(* IEC 61131-3 sources: Industry-PLC-LLM/data/PLCBEAD_repo/PLCBEAD_PLCEmbed-main/PLC-BEAD/Source/PLC_Programs (part 13) *)

(* ---- TN_SC_AREA_RESTORE.ST ---- *)
TYPE
  bya_TN_CHAR:       	ARRAY [0..1919] OF BYTE;
  bya_TN_BACKUP:     	ARRAY [0..1919] OF BYTE;
  bya_TN_COLOR:      	ARRAY [0..1919] OF BYTE;
  bya_TN_Line_Update:	ARRAY [0..23]   OF BOOL;

  us_TN_SCREEN :
  STRUCT
		bya_CHAR:			bya_TN_CHAR;
		bya_COLOR:			bya_TN_COLOR;
		bya_BACKUP:			bya_TN_BACKUP;
		bya_Line_Update:	bya_TN_Line_Update;

		by_Input_Exten_Code:    BYTE;
		by_Input_ASCII_Code:    BYTE;
		bo_Input_ASCII_IsNum:   BOOL;
		in_Page_Number:        	INT;                (* aktive Seiten-Nr.              *)
		in_Cursor_X:           	INT;                (* Cursor X-Position              *)
		in_Cursor_Y:           	INT;                (* Cursor Y-Position              *)
		in_EOS_Offset:         	INT;                (* End of String Offset           *)
		by_Clear_Screen_Attr:  	BYTE;               (* Clear-Screen Attr              *)
		bo_Clear_Screen:       	BOOL;               (* Clear-Screen ausl�sen          *)
		bo_Modal_Dialog:       	BOOL;               (* Modaler Dialog ist aktiv       *)
		bo_Menue_Bar_Dialog:   	BOOL;               (* Menue Dialog ist aktiv         *)

  END_STRUCT;
END_TYPE

FUNCTION TN_SC_XY2_ERROR:BOOL

	VAR_INPUT
		X1 :	INT;
		Y1 :	INT;
		X2 :	INT;
		Y2 :	INT;
	END_VAR

	TN_SC_XY2_ERROR := Y1 < 0 OR X1 < 0 OR Y2 < 0 OR X2 < 0 OR Y1 > 23 OR X1 > 79 OR Y2 > 23 OR X2 > 79;

END_FUNCTION

FUNCTION _BYTE_TO_INT:INT
	VAR_INPUT
		IN :	BYTE;
	END_VAR

	_BYTE_TO_INT := USINT_TO_INT(BYTE_TO_USINT(IN));
END_FUNCTION

FUNCTION_BLOCK TN_SC_AREA_RESTORE_Block

  VAR
    in_Offset_1 :	INT;
    in_Offset_2 :	INT;
    in_Y :	INT;
    in_X :	INT;
    in_Y1 :	INT;
    in_X1 :	INT;
    in_Y2 :	INT;
    in_X2 :	INT;
  END_VAR

  VAR_IN_OUT
    Xus_TN_SCREEN :	us_TN_SCREEN;
  END_VAR

  IF Xus_TN_SCREEN.bya_BACKUP[0] > BYTE#00 THEN

    in_X1 := _BYTE_TO_INT(Xus_TN_SCREEN.bya_BACKUP[1]);
    in_Y1 := _BYTE_TO_INT(Xus_TN_SCREEN.bya_BACKUP[2]);
    in_X2 := _BYTE_TO_INT(Xus_TN_SCREEN.bya_BACKUP[3]);
    in_Y2 := _BYTE_TO_INT(Xus_TN_SCREEN.bya_BACKUP[4]);

    IF TN_SC_XY2_ERROR(in_X1,in_Y1,in_X2,in_Y2) THEN RETURN; END_IF;
    in_Offset_2 := 5;

    FOR in_Y := in_Y1 TO in_Y2 DO

      Xus_TN_SCREEN.bya_Line_Update[in_Y] := TRUE;
      in_Offset_1 := (in_Y * 80) + in_X1;

      FOR in_X := in_X1 TO in_X2 DO

        Xus_TN_SCREEN.bya_CHAR[in_Offset_1] := Xus_TN_SCREEN.bya_BACKUP[in_Offset_2];
        in_Offset_2 := in_Offset_2 + INT#01;

        Xus_TN_SCREEN.bya_COLOR[in_Offset_1] := Xus_TN_SCREEN.bya_BACKUP[in_Offset_2];
        in_Offset_2 := in_Offset_2 + INT#01;
        in_Offset_1 := in_Offset_1 + INT#01;

      END_FOR;

    END_FOR;

    Xus_TN_SCREEN.bya_BACKUP[0] := BYTE#00;
  END_IF;

END_FUNCTION_BLOCK

PROGRAM program0
	VAR
		Xus_TN_SCREEN :	us_TN_SCREEN;

		func_block : TN_SC_AREA_RESTORE_Block;
	END_VAR
	func_block.Xus_TN_SCREEN := Xus_TN_SCREEN;

	func_block();
	Xus_TN_SCREEN  := func_block.Xus_TN_SCREEN;
END_PROGRAM

CONFIGURATION Config0
	RESOURCE Res0 ON PLC
		TASK task0(INTERVAL := T#20ms,PRIORITY := 0);
		PROGRAM instance0 WITH task0 : program0;
	END_RESOURCE
END_CONFIGURATION

(* ---- TN_SC_AREA_SAVE.ST ---- *)
TYPE
  bya_TN_CHAR:       	ARRAY [0..1919] OF BYTE;
  bya_TN_BACKUP:     	ARRAY [0..1919] OF BYTE;
  bya_TN_COLOR:      	ARRAY [0..1919] OF BYTE;
  bya_TN_Line_Update:	ARRAY [0..23]   OF BOOL;

  us_TN_SCREEN :
  STRUCT
		bya_CHAR:			bya_TN_CHAR;
		bya_COLOR:			bya_TN_COLOR;
		bya_BACKUP:			bya_TN_BACKUP;
		bya_Line_Update:	bya_TN_Line_Update;

		by_Input_Exten_Code:    BYTE;
		by_Input_ASCII_Code:    BYTE;
		bo_Input_ASCII_IsNum:   BOOL;
		in_Page_Number:        	INT;                (* aktive Seiten-Nr.              *)
		in_Cursor_X:           	INT;                (* Cursor X-Position              *)
		in_Cursor_Y:           	INT;                (* Cursor Y-Position              *)
		in_EOS_Offset:         	INT;                (* End of String Offset           *)
		by_Clear_Screen_Attr:  	BYTE;               (* Clear-Screen Attr              *)
		bo_Clear_Screen:       	BOOL;               (* Clear-Screen ausl�sen          *)
		bo_Modal_Dialog:       	BOOL;               (* Modaler Dialog ist aktiv       *)
		bo_Menue_Bar_Dialog:   	BOOL;               (* Menue Dialog ist aktiv         *)

  END_STRUCT;
END_TYPE

FUNCTION TN_SC_XY2_ERROR:BOOL

	VAR_INPUT
		X1 :	INT;
		Y1 :	INT;
		X2 :	INT;
		Y2 :	INT;
	END_VAR

	TN_SC_XY2_ERROR := Y1 < 0 OR X1 < 0 OR Y2 < 0 OR X2 < 0 OR Y1 > 23 OR X1 > 79 OR Y2 > 23 OR X2 > 79;

END_FUNCTION

FUNCTION_BLOCK TN_SC_AREA_SAVE_Block

	VAR
		in_Offset_1 :	INT;
		in_Offset_2 :	INT;
		in_Y :	INT;
		in_X :	INT;
	END_VAR

	VAR_INPUT
		Iin_Y1 :	INT;
		Iin_X1 :	INT;
		Iin_Y2 :	INT;
		Iin_X2 :	INT;
	END_VAR

	VAR_IN_OUT
		Xus_TN_SCREEN :	us_TN_SCREEN;
	END_VAR

	IF TN_SC_XY2_ERROR(Iin_X1,Iin_Y1,Iin_X2,Iin_Y2) THEN RETURN; END_IF;

	Xus_TN_SCREEN.bya_BACKUP[0] := BYTE#1;
	Xus_TN_SCREEN.bya_BACKUP[1] := INT_TO_BYTE(Iin_X1);
	Xus_TN_SCREEN.bya_BACKUP[2] := INT_TO_BYTE(Iin_Y1);
	Xus_TN_SCREEN.bya_BACKUP[3] := INT_TO_BYTE(Iin_X2);
	Xus_TN_SCREEN.bya_BACKUP[4] := INT_TO_BYTE(Iin_Y2);

	in_Offset_2 := 5;
	FOR in_Y := Iin_Y1 TO Iin_Y2 DO

	in_Offset_1 := (in_Y * 80) + Iin_X1;
	FOR in_X := Iin_X1 TO Iin_X2 DO

		Xus_TN_SCREEN.bya_BACKUP[in_Offset_2] := Xus_TN_SCREEN.bya_CHAR[in_Offset_1];
		in_Offset_2 := in_Offset_2 + INT#01;
		Xus_TN_SCREEN.bya_BACKUP[in_Offset_2] := Xus_TN_SCREEN.bya_COLOR[in_Offset_1];
		in_Offset_2 := in_Offset_2 + INT#01;
		in_Offset_1 := in_Offset_1 + INT#01;

	END_FOR;
	END_FOR;

END_FUNCTION_BLOCK

PROGRAM program0
	VAR
		Iin_Y1 :	INT;
		Iin_X1 :	INT;
		Iin_Y2 :	INT;
		Iin_X2 :	INT;
		Xus_TN_SCREEN :	us_TN_SCREEN;

		func_block : TN_SC_AREA_SAVE_Block;
	END_VAR
	func_block.Iin_X1 := Iin_X1;
	func_block.Iin_Y1 := Iin_Y1;
	func_block.Iin_X2 := Iin_X2;
	func_block.Iin_Y2 := Iin_Y2;
	func_block.Xus_TN_SCREEN := Xus_TN_SCREEN;

	func_block();
	Xus_TN_SCREEN  := func_block.Xus_TN_SCREEN;
END_PROGRAM

CONFIGURATION Config0
	RESOURCE Res0 ON PLC
		TASK task0(INTERVAL := T#20ms,PRIORITY := 0);
		PROGRAM instance0 WITH task0 : program0;
	END_RESOURCE
END_CONFIGURATION

(* ---- TN_SC_BOX.ST ---- *)
TYPE
  bya_TN_CHAR:       	ARRAY [0..1919] OF BYTE;
  bya_TN_BACKUP:     	ARRAY [0..1919] OF BYTE;
  bya_TN_COLOR:      	ARRAY [0..1919] OF BYTE;
  bya_TN_Line_Update:	ARRAY [0..23]   OF BOOL;

  us_TN_SCREEN :
  STRUCT
		bya_CHAR:			bya_TN_CHAR;
		bya_COLOR:			bya_TN_COLOR;
		bya_BACKUP:			bya_TN_BACKUP;
		bya_Line_Update:	bya_TN_Line_Update;

		by_Input_Exten_Code:    BYTE;
		by_Input_ASCII_Code:    BYTE;
		bo_Input_ASCII_IsNum:   BOOL;
		in_Page_Number:        	INT;                (* aktive Seiten-Nr.              *)
		in_Cursor_X:           	INT;                (* Cursor X-Position              *)
		in_Cursor_Y:           	INT;                (* Cursor Y-Position              *)
		in_EOS_Offset:         	INT;                (* End of String Offset           *)
		by_Clear_Screen_Attr:  	BYTE;               (* Clear-Screen Attr              *)
		bo_Clear_Screen:       	BOOL;               (* Clear-Screen ausl�sen          *)
		bo_Modal_Dialog:       	BOOL;               (* Modaler Dialog ist aktiv       *)
		bo_Menue_Bar_Dialog:   	BOOL;               (* Menue Dialog ist aktiv         *)

  END_STRUCT;
END_TYPE

FUNCTION TN_SC_XY2_ERROR:BOOL

	VAR_INPUT
		X1 :	INT;
		Y1 :	INT;
		X2 :	INT;
		Y2 :	INT;
	END_VAR

	TN_SC_XY2_ERROR := Y1 < 0 OR X1 < 0 OR Y2 < 0 OR X2 < 0 OR Y1 > 23 OR X1 > 79 OR Y2 > 23 OR X2 > 79;

END_FUNCTION

FUNCTION_BLOCK TN_SC_FILL_Block

	VAR
		in_X :	INT;
		in_Y :	INT;
		in_Offset :	INT;
	END_VAR

	VAR_INPUT
		Iin_Y1 :	INT;
		Iin_X1 :	INT;
		Iin_Y2 :	INT;
		Iin_X2 :	INT;
		Iby_CHAR :	BYTE;
		Iby_Attr :	BYTE;
	END_VAR

	VAR_IN_OUT
		Xus_TN_SCREEN :	us_TN_SCREEN;
	END_VAR

	IF TN_SC_XY2_ERROR(Iin_X1,Iin_Y1,Iin_X2,Iin_Y2) THEN RETURN; END_IF;

	FOR in_Y := Iin_Y1 TO Iin_Y2 DO
	Xus_TN_SCREEN.bya_Line_Update[in_Y] := TRUE;
	in_Offset := (in_Y * 80) + Iin_X1;
	FOR in_X := Iin_X1 TO Iin_X2 DO
		Xus_TN_SCREEN.bya_CHAR[in_Offset]  := Iby_CHAR;
		Xus_TN_SCREEN.bya_COLOR[in_Offset] := Iby_Attr;
		in_Offset := in_Offset + 1;
	END_FOR;
	END_FOR;

END_FUNCTION_BLOCK

FUNCTION_BLOCK TN_SC_BOX_Block

  VAR
    FB_TN_SC_FILL :	TN_SC_FILL_Block;
  END_VAR

  VAR
    by_BorderChar_L_T :	BYTE;
    by_BorderChar_T :	BYTE;
    by_BorderChar_B :	BYTE;
    by_BorderChar_R_T :	BYTE;
    by_BorderChar_L :	BYTE;
    by_BorderChar_R :	BYTE;
    by_BorderChar_L_B :	BYTE;
    by_BorderChar_R_B :	BYTE;
    in_Y :	INT;
    in_X :	INT;
    in_Border_Offset :	INT;
    in_Offset_1 :	INT;
    in_Offset_2 :	INT;
  END_VAR

  VAR_INPUT
    Iin_Y1 :	INT;
    Iin_X1 :	INT;
    Iin_Y2 :	INT;
    Iin_X2 :	INT;
    Iby_FILL :	BYTE;
    Iby_ATTR :	BYTE;
    Iin_BORDER :	INT;
  END_VAR

  VAR_IN_OUT
    Xus_TN_SCREEN :	us_TN_SCREEN;
  END_VAR

  IF TN_SC_XY2_ERROR(Iin_X1,Iin_Y1,Iin_X2,Iin_Y2) THEN RETURN; END_IF;

  CASE Iin_Border OF
  0:
    in_Border_Offset := 0;

  1:
    by_BorderChar_L_T := BYTE#218;
    by_BorderChar_T   := BYTE#196;
    by_BorderChar_R_T := BYTE#191;
    by_BorderChar_L   := BYTE#179;
    by_BorderChar_R   := BYTE#179;
    by_BorderChar_B   := BYTE#196;
    by_BorderChar_L_B := BYTE#217;
    by_BorderChar_R_B := BYTE#192;
    in_Border_Offset  := 1;

  2:
    by_BorderChar_L_T := BYTE#201;
    by_BorderChar_T   := BYTE#205;
    by_BorderChar_R_T := BYTE#187;
    by_BorderChar_L   := BYTE#186;
    by_BorderChar_R   := BYTE#186;
    by_BorderChar_B   := BYTE#205;
    by_BorderChar_L_B := BYTE#188;
    by_BorderChar_R_B := BYTE#200;
    in_Border_Offset  := 1;

  ELSE
    by_BorderChar_L_T := BYTE#32;
    by_BorderChar_T   := BYTE#32;
    by_BorderChar_R_T := BYTE#32;
    by_BorderChar_L   := BYTE#32;
    by_BorderChar_R   := BYTE#32;
    by_BorderChar_B   := BYTE#32;
    by_BorderChar_L_B := BYTE#32;
    by_BorderChar_R_B := BYTE#32;
    in_Border_Offset  := 1;

  END_CASE;

  IF Iby_FILL > BYTE#0 THEN

    FB_TN_SC_FILL.Iin_Y1			:= Iin_Y1 + in_Border_Offset;
    FB_TN_SC_FILL.Iin_X1			:= Iin_X1 + in_Border_Offset;
    FB_TN_SC_FILL.Iin_Y2			:= Iin_Y2 - in_Border_Offset;
    FB_TN_SC_FILL.Iin_X2			:= Iin_X2 - in_Border_Offset;
    FB_TN_SC_FILL.Iby_CHAR		:= Iby_FILL;
    FB_TN_SC_FILL.Iby_Attr		:= Iby_ATTR;
    FB_TN_SC_FILL.Xus_TN_SCREEN := Xus_TN_SCREEN;
    FB_TN_SC_FILL();
    Xus_TN_SCREEN := FB_TN_SC_FILL.Xus_TN_SCREEN;

  END_IF;

  IF Iin_BORDER = 0 THEN RETURN; END_IF;

  in_Offset_1 := (Iin_Y1 * 80) + Iin_X1;
  in_Offset_2 := (Iin_Y1 * 80) + Iin_X2;

  FOR in_Y := Iin_Y1 TO Iin_Y2 DO

    Xus_TN_SCREEN.bya_Line_Update[in_Y] := TRUE;

    Xus_TN_SCREEN.bya_CHAR[in_Offset_1]  := by_BorderChar_L;
    Xus_TN_SCREEN.bya_COLOR[in_Offset_1] := Iby_Attr;

    Xus_TN_SCREEN.bya_CHAR[in_Offset_2]  := by_BorderChar_R;
    Xus_TN_SCREEN.bya_COLOR[in_Offset_2] := Iby_Attr;

    in_Offset_1 := in_Offset_1 + 80;
    in_Offset_2 := in_Offset_2 + 80;

  END_FOR;

  in_Offset_1 := (Iin_Y1 * 80) + Iin_X1;
  in_Offset_2 := (Iin_Y2 * 80) + Iin_X1;

  FOR in_X := Iin_X1 TO Iin_X2 DO

    Xus_TN_SCREEN.bya_CHAR[in_Offset_1]  := by_BorderChar_T;
    Xus_TN_SCREEN.bya_COLOR[in_Offset_1] := Iby_Attr;

    Xus_TN_SCREEN.bya_CHAR[in_Offset_2]  := by_BorderChar_B;
    Xus_TN_SCREEN.bya_COLOR[in_Offset_2] := Iby_Attr;

    in_Offset_1 := in_Offset_1 + INT#1;
    in_Offset_2 := in_Offset_2 + INT#1;

  END_FOR;

  in_Offset_1 := (Iin_Y1 * 80) + Iin_X1;
  Xus_TN_SCREEN.bya_CHAR[in_Offset_1]  := by_BorderChar_L_T;
  Xus_TN_SCREEN.bya_COLOR[in_Offset_1] := Iby_Attr;

  in_Offset_1 := (Iin_Y1 * 80) + Iin_X2;
  Xus_TN_SCREEN.bya_CHAR[in_Offset_1]  := by_BorderChar_R_T;
  Xus_TN_SCREEN.bya_COLOR[in_Offset_1] := Iby_Attr;

  in_Offset_1 := (Iin_Y2 * 80) + Iin_X1;
  Xus_TN_SCREEN.bya_CHAR[in_Offset_1]  := by_BorderChar_R_B;
  Xus_TN_SCREEN.bya_COLOR[in_Offset_1] := Iby_Attr;

  in_Offset_1 := (Iin_Y2 * 80) + Iin_X2;
  Xus_TN_SCREEN.bya_CHAR[in_Offset_1]  := by_BorderChar_L_B;
  Xus_TN_SCREEN.bya_COLOR[in_Offset_1] := Iby_Attr;

END_FUNCTION_BLOCK

PROGRAM program0
	VAR
		Iin_Y1 :	INT;
    Iin_X1 :	INT;
    Iin_Y2 :	INT;
    Iin_X2 :	INT;
    Iby_FILL :	BYTE;
    Iby_ATTR :	BYTE;
    Iin_BORDER :	INT;
		Xus_TN_SCREEN :	us_TN_SCREEN;

		func_block : TN_SC_BOX_Block;
	END_VAR
  func_block.Iin_X1 := Iin_X1;
  func_block.Iin_Y1 := Iin_Y1;
  func_block.Iin_X2 := Iin_X2;
  func_block.Iin_Y2 := Iin_Y2;
  func_block.Iby_FILL := Iby_FILL;
  func_block.Iby_ATTR := Iby_ATTR;
  func_block.Iin_BORDER := Iin_BORDER;
  func_block.Xus_TN_SCREEN := Xus_TN_SCREEN;

	func_block();
	Xus_TN_SCREEN  := func_block.Xus_TN_SCREEN;
END_PROGRAM

CONFIGURATION Config0
	RESOURCE Res0 ON PLC
		TASK task0(INTERVAL := T#20ms,PRIORITY := 0);
		PROGRAM instance0 WITH task0 : program0;
	END_RESOURCE
END_CONFIGURATION

(* ---- TN_SC_FILL.ST ---- *)
TYPE
  bya_TN_CHAR:       	ARRAY [0..1919] OF BYTE;
  bya_TN_BACKUP:     	ARRAY [0..1919] OF BYTE;
  bya_TN_COLOR:      	ARRAY [0..1919] OF BYTE;
  bya_TN_Line_Update:	ARRAY [0..23]   OF BOOL;

  us_TN_SCREEN :
  STRUCT
		bya_CHAR:			bya_TN_CHAR;
		bya_COLOR:			bya_TN_COLOR;
		bya_BACKUP:			bya_TN_BACKUP;
		bya_Line_Update:	bya_TN_Line_Update;

		by_Input_Exten_Code:    BYTE;
		by_Input_ASCII_Code:    BYTE;
		bo_Input_ASCII_IsNum:   BOOL;
		in_Page_Number:        	INT;                (* aktive Seiten-Nr.              *)
		in_Cursor_X:           	INT;                (* Cursor X-Position              *)
		in_Cursor_Y:           	INT;                (* Cursor Y-Position              *)
		in_EOS_Offset:         	INT;                (* End of String Offset           *)
		by_Clear_Screen_Attr:  	BYTE;               (* Clear-Screen Attr              *)
		bo_Clear_Screen:       	BOOL;               (* Clear-Screen ausl�sen          *)
		bo_Modal_Dialog:       	BOOL;               (* Modaler Dialog ist aktiv       *)
		bo_Menue_Bar_Dialog:   	BOOL;               (* Menue Dialog ist aktiv         *)

  END_STRUCT;
END_TYPE

FUNCTION TN_SC_XY2_ERROR:BOOL

	VAR_INPUT
		X1 :	INT;
		Y1 :	INT;
		X2 :	INT;
		Y2 :	INT;
	END_VAR

	TN_SC_XY2_ERROR := Y1 < 0 OR X1 < 0 OR Y2 < 0 OR X2 < 0 OR Y1 > 23 OR X1 > 79 OR Y2 > 23 OR X2 > 79;

END_FUNCTION

FUNCTION_BLOCK TN_SC_FILL_Block

	VAR
		in_X :	INT;
		in_Y :	INT;
		in_Offset :	INT;
	END_VAR

	VAR_INPUT
		Iin_Y1 :	INT;
		Iin_X1 :	INT;
		Iin_Y2 :	INT;
		Iin_X2 :	INT;
		Iby_CHAR :	BYTE;
		Iby_Attr :	BYTE;
	END_VAR

	VAR_IN_OUT
		Xus_TN_SCREEN :	us_TN_SCREEN;
	END_VAR

	IF TN_SC_XY2_ERROR(Iin_X1,Iin_Y1,Iin_X2,Iin_Y2) THEN RETURN; END_IF;

	FOR in_Y := Iin_Y1 TO Iin_Y2 DO
	Xus_TN_SCREEN.bya_Line_Update[in_Y] := TRUE;
	in_Offset := (in_Y * 80) + Iin_X1;
	FOR in_X := Iin_X1 TO Iin_X2 DO
		Xus_TN_SCREEN.bya_CHAR[in_Offset]  := Iby_CHAR;
		Xus_TN_SCREEN.bya_COLOR[in_Offset] := Iby_Attr;
		in_Offset := in_Offset + 1;
	END_FOR;
	END_FOR;

END_FUNCTION_BLOCK

PROGRAM program0
	VAR
		Iin_Y1 :	INT;
		Iin_X1 :	INT;
		Iin_Y2 :	INT;
		Iin_X2 :	INT;
		Iby_CHAR :	BYTE;
		Iby_Attr :	BYTE;
		Xus_TN_SCREEN :	us_TN_SCREEN;

		func_block : TN_SC_FILL_Block;
	END_VAR
	func_block.Iin_X1 := Iin_X1;
	func_block.Iin_Y1 := Iin_Y1;
  	func_block.Iin_X2 := Iin_X2;
	func_block.Iin_Y2 := Iin_Y2;
  	func_block.Iby_CHAR := Iby_CHAR;
	func_block.Iby_Attr := Iby_Attr;
	func_block.Xus_TN_SCREEN := Xus_TN_SCREEN;

	func_block();
	Xus_TN_SCREEN  := func_block.Xus_TN_SCREEN;
END_PROGRAM

CONFIGURATION Config0
	RESOURCE Res0 ON PLC
		TASK task0(INTERVAL := T#20ms,PRIORITY := 0);
		PROGRAM instance0 WITH task0 : program0;
	END_RESOURCE
END_CONFIGURATION

(* ---- TN_SC_LINE.ST ---- *)
TYPE
  bya_TN_CHAR:       	ARRAY [0..1919] OF BYTE;
  bya_TN_BACKUP:     	ARRAY [0..1919] OF BYTE;
  bya_TN_COLOR:      	ARRAY [0..1919] OF BYTE;
  bya_TN_Line_Update:	ARRAY [0..23]   OF BOOL;

  us_TN_SCREEN :
  STRUCT
		bya_CHAR:			bya_TN_CHAR;
		bya_COLOR:			bya_TN_COLOR;
		bya_BACKUP:			bya_TN_BACKUP;
		bya_Line_Update:	bya_TN_Line_Update;

		by_Input_Exten_Code:    BYTE;
		by_Input_ASCII_Code:    BYTE;
		bo_Input_ASCII_IsNum:   BOOL;
		in_Page_Number:        	INT;                (* aktive Seiten-Nr.              *)
		in_Cursor_X:           	INT;                (* Cursor X-Position              *)
		in_Cursor_Y:           	INT;                (* Cursor Y-Position              *)
		in_EOS_Offset:         	INT;                (* End of String Offset           *)
		by_Clear_Screen_Attr:  	BYTE;               (* Clear-Screen Attr              *)
		bo_Clear_Screen:       	BOOL;               (* Clear-Screen ausl�sen          *)
		bo_Modal_Dialog:       	BOOL;               (* Modaler Dialog ist aktiv       *)
		bo_Menue_Bar_Dialog:   	BOOL;               (* Menue Dialog ist aktiv         *)

  END_STRUCT;
END_TYPE

FUNCTION TN_SC_XY2_ERROR:BOOL

	VAR_INPUT
		X1 :	INT;
		Y1 :	INT;
		X2 :	INT;
		Y2 :	INT;
	END_VAR

	TN_SC_XY2_ERROR := Y1 < 0 OR X1 < 0 OR Y2 < 0 OR X2 < 0 OR Y1 > 23 OR X1 > 79 OR Y2 > 23 OR X2 > 79;

END_FUNCTION

FUNCTION_BLOCK TN_SC_LINE_Block

  VAR
    by_Connect_Left_Char :	BYTE;
    by_Connect_Right_Char :	BYTE;
    by_Connect_Top_Char :	BYTE;
    by_Connect_Bottom_Char :	BYTE;
    by_Connect_Cruz_Char :	BYTE;
    by_Vertikal_Line_Char :	BYTE;
    by_Horzontal_Line_Char :	BYTE;
    by_old_Char :	BYTE;
    in_Offset_1 :	INT;
    in_ROW_Index :	INT;
    in_COL_Index :	INT;
    by_Char :	BYTE;
  END_VAR

  VAR_INPUT
    Iin_X1 :	INT;
    Iin_Y1 :	INT;
    Iin_X2 :	INT;
    Iin_Y2 :	INT;
    Iby_ATTR :	BYTE;
    Iby_BORDER :	BYTE;
  END_VAR

  VAR_IN_OUT
    Xus_TN_SCREEN :	us_TN_SCREEN;
  END_VAR

  IF TN_SC_XY2_ERROR(Iin_X1,Iin_Y1,Iin_X2,Iin_Y2) THEN RETURN; END_IF;

  IF Iby_Border = BYTE#01 THEN

    by_Connect_Top_Char    := BYTE#16#C2;
    by_Connect_Bottom_Char := BYTE#16#C1;
    by_Connect_Left_Char   := BYTE#16#C3;
    by_Connect_Right_Char  := BYTE#16#B4;
    by_Horzontal_Line_Char := BYTE#16#C4;
    by_Vertikal_Line_Char  := BYTE#16#B3;
    by_Connect_Cruz_Char   := BYTE#16#C5;

  ELSIF Iby_Border = BYTE#02 THEN

    by_Connect_Top_Char    := BYTE#16#CB;
    by_Connect_Bottom_Char := BYTE#16#CA;
    by_Connect_Left_Char   := BYTE#16#CC;
    by_Connect_Right_Char  := BYTE#16#B9;
    by_Horzontal_Line_Char := BYTE#16#CD;
    by_Vertikal_Line_Char  := BYTE#16#BA;
    by_Connect_Cruz_Char   := BYTE#16#CE;

  ELSE
    by_Connect_Top_Char    := Iby_Border;
    by_Connect_Bottom_Char := Iby_Border;
    by_Connect_Left_Char   := Iby_Border;
    by_Connect_Right_Char  := Iby_Border;
    by_Horzontal_Line_Char := Iby_Border;
    by_Vertikal_Line_Char  := Iby_Border;
    by_Connect_Cruz_Char   := Iby_Border;

  END_IF;

  IF Iin_X1 = Iin_X2 THEN

    in_Offset_1 := (Iin_Y1 * 80) + Iin_X1;

    FOR in_ROW_Index := Iin_Y1 TO Iin_Y2 DO

      by_old_Char := Xus_TN_SCREEN.bya_CHAR[in_Offset_1];

      by_Char := by_Vertikal_Line_Char;

      IF by_old_Char = by_Horzontal_Line_Char THEN

        IF in_ROW_Index = Iin_Y1 THEN
          by_Char := by_Connect_Top_Char;

        ELSIF in_ROW_Index = Iin_Y2 THEN
          by_Char := by_Connect_Bottom_Char;

        ELSE
          by_Char := by_Connect_Cruz_Char;
        END_IF;

      END_IF;

      Xus_TN_SCREEN.bya_Line_Update[in_ROW_Index] := TRUE;

      Xus_TN_SCREEN.bya_CHAR[in_Offset_1]  := by_Char;
      Xus_TN_SCREEN.bya_COLOR[in_Offset_1] := Iby_Attr;

      in_Offset_1 := in_Offset_1 + 80;

    END_FOR;

  ELSIF Iin_Y1 = Iin_Y2 THEN

    Xus_TN_SCREEN.bya_Line_Update[Iin_Y1] := TRUE;

    in_Offset_1 := (Iin_Y1 * 80) + Iin_X1;

    FOR in_COL_Index := Iin_X1 TO Iin_X2 DO

      by_old_Char := Xus_TN_SCREEN.bya_CHAR[in_Offset_1];

      by_Char := by_Horzontal_Line_Char;

      IF by_old_Char = by_Vertikal_Line_Char THEN

        IF in_COL_Index = Iin_X1 THEN
          by_Char := by_Connect_Left_Char;

        ELSIF in_COL_Index = Iin_X2 THEN
          by_Char := by_Connect_Right_Char;

        ELSE
          by_Char := by_Connect_Cruz_Char;
        END_IF;

      END_IF;

      Xus_TN_SCREEN.bya_CHAR[in_Offset_1]  := by_Char;
      Xus_TN_SCREEN.bya_COLOR[in_Offset_1] := Iby_Attr;

      in_Offset_1 := in_Offset_1 + 1;

    END_FOR;
  END_IF;

END_FUNCTION_BLOCK

PROGRAM program0
	VAR
    Iin_X1 :	INT;
    Iin_Y1 :	INT;
    Iin_X2 :	INT;
    Iin_Y2 :	INT;
    Iby_ATTR :	BYTE;
    Iby_BORDER :	BYTE;
    Xus_TN_SCREEN :	us_TN_SCREEN;

    func_block : TN_SC_LINE_Block;
	END_VAR
	func_block.Iin_X1 := Iin_X1;
	func_block.Iin_Y1 := Iin_Y1;
  func_block.Iin_X2 := Iin_X2;
	func_block.Iin_Y2 := Iin_Y2;
  func_block.Iby_ATTR := Iby_ATTR;
	func_block.Iby_BORDER := Iby_BORDER;
	func_block.Xus_TN_SCREEN := Xus_TN_SCREEN;

	func_block();
	Xus_TN_SCREEN  := func_block.Xus_TN_SCREEN;
END_PROGRAM

CONFIGURATION Config0
	RESOURCE Res0 ON PLC
		TASK task0(INTERVAL := T#20ms,PRIORITY := 0);
		PROGRAM instance0 WITH task0 : program0;
	END_RESOURCE
END_CONFIGURATION

(* ---- TN_SC_READ_ATTR.ST ---- *)
TYPE
  bya_TN_CHAR:       	ARRAY [0..1919] OF BYTE;
  bya_TN_BACKUP:     	ARRAY [0..1919] OF BYTE;
  bya_TN_COLOR:      	ARRAY [0..1919] OF BYTE;
  bya_TN_Line_Update:	ARRAY [0..23]   OF BOOL;

  us_TN_SCREEN :
  STRUCT
		bya_CHAR:			bya_TN_CHAR;
		bya_COLOR:			bya_TN_COLOR;
		bya_BACKUP:			bya_TN_BACKUP;
		bya_Line_Update:	bya_TN_Line_Update;

		by_Input_Exten_Code:    BYTE;
		by_Input_ASCII_Code:    BYTE;
		bo_Input_ASCII_IsNum:   BOOL;
		in_Page_Number:        	INT;                (* aktive Seiten-Nr.              *)
		in_Cursor_X:           	INT;                (* Cursor X-Position              *)
		in_Cursor_Y:           	INT;                (* Cursor Y-Position              *)
		in_EOS_Offset:         	INT;                (* End of String Offset           *)
		by_Clear_Screen_Attr:  	BYTE;               (* Clear-Screen Attr              *)
		bo_Clear_Screen:       	BOOL;               (* Clear-Screen ausl�sen          *)
		bo_Modal_Dialog:       	BOOL;               (* Modaler Dialog ist aktiv       *)
		bo_Menue_Bar_Dialog:   	BOOL;               (* Menue Dialog ist aktiv         *)

  END_STRUCT;
END_TYPE

FUNCTION TN_SC_XY_ERROR:BOOL

	VAR_INPUT
		X :	INT;
		Y :	INT;
	END_VAR

	TN_SC_XY_ERROR := Y < 0 OR X < 0 OR Y > 23 OR X > 79;

END_FUNCTION

FUNCTION_BLOCK TN_SC_READ_ATTR_Block

	VAR
		in_Offset :	INT;
	END_VAR

	VAR_INPUT
		Iin_Y :	INT;
		Iin_X :	INT;
	END_VAR

	VAR_OUTPUT
		Oby_ATTR :	BYTE;
	END_VAR

	VAR_IN_OUT
		Xus_TN_SCREEN :	us_TN_SCREEN;
	END_VAR

	IF TN_SC_XY_ERROR(Iin_X,Iin_Y) THEN RETURN; END_IF;
	in_Offset := (Iin_Y * 80) + Iin_X;
	Oby_ATTR := Xus_TN_SCREEN.bya_COLOR[in_Offset];

END_FUNCTION_BLOCK

PROGRAM program0
	VAR
		Iin_Y :	INT;
		Iin_X :	INT;
		Xus_TN_SCREEN :	us_TN_SCREEN;
		Oby_ATTR :	BYTE;

		func_block : TN_SC_READ_ATTR_Block;
	END_VAR
	func_block.Iin_Y := Iin_Y;
	func_block.Iin_X := Iin_X;
	func_block.Xus_TN_SCREEN := Xus_TN_SCREEN;

	func_block();
	Xus_TN_SCREEN  := func_block.Xus_TN_SCREEN;
	Oby_ATTR  := func_block.Oby_ATTR;
END_PROGRAM

CONFIGURATION Config0
	RESOURCE Res0 ON PLC
		TASK task0(INTERVAL := T#20ms,PRIORITY := 0);
		PROGRAM instance0 WITH task0 : program0;
	END_RESOURCE
END_CONFIGURATION

(* ---- TN_SC_READ_CHAR.ST ---- *)
TYPE
  bya_TN_CHAR:       	ARRAY [0..1919] OF BYTE;
  bya_TN_BACKUP:     	ARRAY [0..1919] OF BYTE;
  bya_TN_COLOR:      	ARRAY [0..1919] OF BYTE;
  bya_TN_Line_Update:	ARRAY [0..23]   OF BOOL;

  us_TN_SCREEN :
  STRUCT
		bya_CHAR:			bya_TN_CHAR;
		bya_COLOR:			bya_TN_COLOR;
		bya_BACKUP:			bya_TN_BACKUP;
		bya_Line_Update:	bya_TN_Line_Update;

		by_Input_Exten_Code:    BYTE;
		by_Input_ASCII_Code:    BYTE;
		bo_Input_ASCII_IsNum:   BOOL;
		in_Page_Number:        	INT;                (* aktive Seiten-Nr.              *)
		in_Cursor_X:           	INT;                (* Cursor X-Position              *)
		in_Cursor_Y:           	INT;                (* Cursor Y-Position              *)
		in_EOS_Offset:         	INT;                (* End of String Offset           *)
		by_Clear_Screen_Attr:  	BYTE;               (* Clear-Screen Attr              *)
		bo_Clear_Screen:       	BOOL;               (* Clear-Screen ausl�sen          *)
		bo_Modal_Dialog:       	BOOL;               (* Modaler Dialog ist aktiv       *)
		bo_Menue_Bar_Dialog:   	BOOL;               (* Menue Dialog ist aktiv         *)

  END_STRUCT;
END_TYPE

FUNCTION TN_SC_XY_ERROR:BOOL

	VAR_INPUT
		X :	INT;
		Y :	INT;
	END_VAR

	TN_SC_XY_ERROR := Y < 0 OR X < 0 OR Y > 23 OR X > 79;

END_FUNCTION

FUNCTION_BLOCK TN_SC_READ_CHAR_Block

	VAR
		in_Offset :	INT;
	END_VAR

	VAR_INPUT
		Iin_Y :	INT;
		Iin_X :	INT;
	END_VAR

	VAR_OUTPUT
		Oby_CHAR :	BYTE;
	END_VAR

	VAR_IN_OUT
		Xus_TN_SCREEN :	us_TN_SCREEN;
	END_VAR

	IF TN_SC_XY_ERROR(Iin_X,Iin_Y) THEN RETURN; END_IF;
	in_Offset := (Iin_Y * 80) + Iin_X;
	Oby_CHAR := Xus_TN_SCREEN.bya_CHAR[in_Offset];

END_FUNCTION_BLOCK

PROGRAM program0
	VAR
		Iin_Y :	INT;
		Iin_X :	INT;
		Xus_TN_SCREEN :	us_TN_SCREEN;
		Oby_CHAR :	BYTE;

		func_block : TN_SC_READ_CHAR_Block;
	END_VAR
	func_block.Iin_Y := Iin_Y;
	func_block.Iin_X := Iin_X;
	func_block.Xus_TN_SCREEN := Xus_TN_SCREEN;

	func_block();
	Xus_TN_SCREEN  := func_block.Xus_TN_SCREEN;
	Oby_CHAR  := func_block.Oby_CHAR;
END_PROGRAM

CONFIGURATION Config0
	RESOURCE Res0 ON PLC
		TASK task0(INTERVAL := T#20ms,PRIORITY := 0);
		PROGRAM instance0 WITH task0 : program0;
	END_RESOURCE
END_CONFIGURATION

(* ---- TN_SC_VIEWPORT.ST ---- *)
TYPE
  bya_TN_CHAR:       	ARRAY [0..1919] OF BYTE;
  bya_TN_BACKUP:     	ARRAY [0..1919] OF BYTE;
  bya_TN_COLOR:      	ARRAY [0..1919] OF BYTE;
  bya_TN_Line_Update:	ARRAY [0..23]   OF BOOL;

  us_TN_SCREEN :
  STRUCT
		bya_CHAR:			bya_TN_CHAR;
		bya_COLOR:			bya_TN_COLOR;
		bya_BACKUP:			bya_TN_BACKUP;
		bya_Line_Update:	bya_TN_Line_Update;

		by_Input_Exten_Code:    BYTE;
		by_Input_ASCII_Code:    BYTE;
		bo_Input_ASCII_IsNum:   BOOL;
		in_Page_Number:        	INT;                (* aktive Seiten-Nr.              *)
		in_Cursor_X:           	INT;                (* Cursor X-Position              *)
		in_Cursor_Y:           	INT;                (* Cursor Y-Position              *)
		in_EOS_Offset:         	INT;                (* End of String Offset           *)
		by_Clear_Screen_Attr:  	BYTE;               (* Clear-Screen Attr              *)
		bo_Clear_Screen:       	BOOL;               (* Clear-Screen ausl�sen          *)
		bo_Modal_Dialog:       	BOOL;               (* Modaler Dialog ist aktiv       *)
		bo_Menue_Bar_Dialog:   	BOOL;               (* Menue Dialog ist aktiv         *)

  END_STRUCT;
END_TYPE

FUNCTION_BLOCK TN_SC_VIEWPORT_Block

  VAR
    FB_TN_SC_WRITE :	TN_SC_WRITE;
    FB_FIX :	FIX;
    FB_TON :	TON;
  END_VAR

  VAR
    in_index :	INT;
    in_Color :	INT;
    by_Attr :	BYTE;
    in_count :	INT;
  END_VAR

  VAR_IN_OUT
    Xus_LOG_VIEWPORT :	us_LOG_VIEWPORT;
    Xus_LOG_CONTROL :	us_LOG_CONTROL_80;
    Xus_TN_SCREEN :	us_TN_SCREEN;
  END_VAR

  VAR_INPUT
    Iin_X :	INT;
    Iin_Y :	INT;
    Iin_Width :	INT;
    Idw_ATTR_1 :	DWORD;
    Idw_ATTR_2 :	DWORD;
    Iti_TIME :	TIME;
  END_VAR

  IF Xus_LOG_VIEWPORT.UPDATE AND FB_TON.Q THEN

    Xus_LOG_VIEWPORT.UPDATE := FALSE;

    FOR in_count := 1 TO Xus_LOG_VIEWPORT.COUNT DO

      in_index := Xus_LOG_VIEWPORT.LINE_ARRAY[in_count];

    in_Color := DWORD_TO_INT(Xus_LOG_CONTROL.MSG_OPTION[in_index] AND DWORD#2#1111);

      CASE in_Color OF
        0..3: by_Attr := BYTE_OF_DWORD(Idw_ATTR_1,INT_TO_BYTE(in_Color));
        4..7: by_Attr := BYTE_OF_DWORD(Idw_ATTR_2,INT_TO_BYTE(in_Color));
      ELSE
      by_Attr := BYTE_OF_DWORD(Idw_ATTR_1,BYTE#0);
      END_CASE;

      FB_FIX.str := Xus_LOG_CONTROL.MSG[in_index];
      FB_FIX.L   := Iin_Width;
      FB_FIX.C   := BYTE#32;
      FB_FIX.M   := INT#00;
      FB_FIX();

      FB_TN_SC_WRITE.Iin_Y			:= Iin_Y + in_count - INT#01;
      FB_TN_SC_WRITE.Iin_X			:= Iin_X;
      FB_TN_SC_WRITE.Iby_ATTR			:= by_Attr;
      FB_TN_SC_WRITE.Ist_STRING		:= FB_FIX.FIX;
      FB_TN_SC_WRITE.Xus_TN_SCREEN	:= Xus_TN_SCREEN;
      FB_TN_SC_WRITE();
      Xus_TN_SCREEN := FB_TN_SC_WRITE.Xus_TN_SCREEN;

    END_FOR;

    FB_TON.IN := FALSE;
    FB_TON.PT := Iti_TIME;
    FB_TON();

  END_IF;

  FB_TON.IN := TRUE;
  FB_TON.PT := Iti_TIME;
  FB_TON();

END_FUNCTION_BLOCK

PROGRAM program0
	VAR
		Xus_LOG_VIEWPORT :	us_LOG_VIEWPORT;
    Xus_LOG_CONTROL :	us_LOG_CONTROL_80;
    Xus_TN_SCREEN :	us_TN_SCREEN;
    Iin_X :	INT;
    Iin_Y :	INT;
    Iin_Width :	INT;
    Idw_ATTR_1 :	DWORD;
    Idw_ATTR_2 :	DWORD;
    Iti_TIME :	TIME;

		func_block : TN_SC_VIEWPORT_Block;
	END_VAR
	func_block.Xus_LOG_VIEWPORT := Xus_LOG_VIEWPORT;
	func_block.Xus_LOG_CONTROL := Xus_LOG_CONTROL;
	func_block.Xus_TN_SCREEN := Xus_TN_SCREEN;
	func_block.Iin_X := Iin_X;
  func_block.Iin_Y := Iin_Y;
	func_block.Iin_Width := Iin_Width;
	func_block.Idw_ATTR_1 := Idw_ATTR_1;
	func_block.Idw_ATTR_2 := Idw_ATTR_2;
  func_block.Iti_TIME := Iti_TIME;

	func_block();
	Xus_LOG_VIEWPORT  := func_block.Xus_LOG_VIEWPORT;
  Xus_LOG_CONTROL  := func_block.Xus_LOG_CONTROL;
  Xus_TN_SCREEN  := func_block.Xus_TN_SCREEN;
END_PROGRAM

CONFIGURATION Config0
	RESOURCE Res0 ON PLC
		TASK task0(INTERVAL := T#20ms,PRIORITY := 0);
		PROGRAM instance0 WITH task0 : program0;
	END_RESOURCE
END_CONFIGURATION

(* ---- TN_SC_WRITE.ST ---- *)
TYPE
  bya_TN_CHAR:       	ARRAY [0..1919] OF BYTE;
  bya_TN_BACKUP:     	ARRAY [0..1919] OF BYTE;
  bya_TN_COLOR:      	ARRAY [0..1919] OF BYTE;
  bya_TN_Line_Update:	ARRAY [0..23]   OF BOOL;

  us_TN_SCREEN :
  STRUCT
		bya_CHAR:			bya_TN_CHAR;
		bya_COLOR:			bya_TN_COLOR;
		bya_BACKUP:			bya_TN_BACKUP;
		bya_Line_Update:	bya_TN_Line_Update;

		by_Input_Exten_Code:    BYTE;
		by_Input_ASCII_Code:    BYTE;
		bo_Input_ASCII_IsNum:   BOOL;
		in_Page_Number:        	INT;                (* aktive Seiten-Nr.              *)
		in_Cursor_X:           	INT;                (* Cursor X-Position              *)
		in_Cursor_Y:           	INT;                (* Cursor Y-Position              *)
		in_EOS_Offset:         	INT;                (* End of String Offset           *)
		by_Clear_Screen_Attr:  	BYTE;               (* Clear-Screen Attr              *)
		bo_Clear_Screen:       	BOOL;               (* Clear-Screen ausl�sen          *)
		bo_Modal_Dialog:       	BOOL;               (* Modaler Dialog ist aktiv       *)
		bo_Menue_Bar_Dialog:   	BOOL;               (* Menue Dialog ist aktiv         *)

  END_STRUCT;
END_TYPE

FUNCTION TN_SC_XY_ERROR:BOOL

	VAR_INPUT
		X :	INT;
		Y :	INT;
	END_VAR

	TN_SC_XY_ERROR := Y < 0 OR X < 0 OR Y > 23 OR X > 79;

END_FUNCTION

FUNCTION_BLOCK TN_SC_WRITE_Block

	VAR
		CODE :	CODE;
	END_VAR

	VAR
		bo_Color :	BOOL;
		in_Offset :	INT;
		in_Char_Index :	INT;
		in_String_Length :	INT;
	END_VAR

	VAR_INPUT
		Iin_Y :	INT;
		Iin_X :	INT;
		Iby_ATTR :	BYTE;
		Ist_STRING :	STRING;
	END_VAR

	VAR_IN_OUT
		Xus_TN_SCREEN :	us_TN_SCREEN;
	END_VAR

	in_String_Length := LEN(Ist_STRING);
	IF TN_SC_XY_ERROR(Iin_X + in_String_Length - 1,Iin_Y) THEN RETURN; END_IF;
	Xus_TN_SCREEN.bya_Line_Update[Iin_Y] := TRUE;
	in_Offset := (Iin_Y * 80) + Iin_X;
	bo_Color := Iby_ATTR <> BYTE#00;

	FOR in_Char_Index := 1 TO in_String_Length DO

	IF bo_Color THEN Xus_TN_SCREEN.bya_COLOR[in_Offset] := Iby_ATTR; END_IF;

	CODE(STR:=Ist_STRING,POS:=in_Char_Index);
	Xus_TN_SCREEN.bya_CHAR[in_Offset] := CODE.CODE;
	in_Offset := in_Offset + INT#1;

	END_FOR;

	Xus_TN_SCREEN.in_EOS_Offset := in_Offset;

END_FUNCTION_BLOCK

PROGRAM program0
	VAR
		Iin_Y :	INT;
		Iin_X :	INT;
		Iby_ATTR :	BYTE;
		Ist_STRING :	STRING;
		Xus_TN_SCREEN :	us_TN_SCREEN;

		func_block : TN_SC_WRITE_Block;
	END_VAR
	func_block.Iin_Y := Iin_Y;
	func_block.Iin_X := Iin_X;
	func_block.Iby_ATTR := Iby_ATTR;
	func_block.Ist_STRING := Ist_STRING;
	func_block.Xus_TN_SCREEN := Xus_TN_SCREEN;

	func_block();
	Xus_TN_SCREEN  := func_block.Xus_TN_SCREEN;

END_PROGRAM

CONFIGURATION Config0
	RESOURCE Res0 ON PLC
		TASK task0(INTERVAL := T#20ms,PRIORITY := 0);
		PROGRAM instance0 WITH task0 : program0;
	END_RESOURCE
END_CONFIGURATION

(* ---- TN_SC_WRITE_ATTR.ST ---- *)
TYPE
  bya_TN_CHAR:       	ARRAY [0..1919] OF BYTE;
  bya_TN_BACKUP:     	ARRAY [0..1919] OF BYTE;
  bya_TN_COLOR:      	ARRAY [0..1919] OF BYTE;
  bya_TN_Line_Update:	ARRAY [0..23]   OF BOOL;

  us_TN_SCREEN :
  STRUCT
		bya_CHAR:			bya_TN_CHAR;
		bya_COLOR:			bya_TN_COLOR;
		bya_BACKUP:			bya_TN_BACKUP;
		bya_Line_Update:	bya_TN_Line_Update;

		by_Input_Exten_Code:    BYTE;
		by_Input_ASCII_Code:    BYTE;
		bo_Input_ASCII_IsNum:   BOOL;
		in_Page_Number:        	INT;                (* aktive Seiten-Nr.              *)
		in_Cursor_X:           	INT;                (* Cursor X-Position              *)
		in_Cursor_Y:           	INT;                (* Cursor Y-Position              *)
		in_EOS_Offset:         	INT;                (* End of String Offset           *)
		by_Clear_Screen_Attr:  	BYTE;               (* Clear-Screen Attr              *)
		bo_Clear_Screen:       	BOOL;               (* Clear-Screen ausl�sen          *)
		bo_Modal_Dialog:       	BOOL;               (* Modaler Dialog ist aktiv       *)
		bo_Menue_Bar_Dialog:   	BOOL;               (* Menue Dialog ist aktiv         *)

  END_STRUCT;
END_TYPE

FUNCTION TN_SC_XY_ERROR:BOOL

	VAR_INPUT
		X :	INT;
		Y :	INT;
	END_VAR

	TN_SC_XY_ERROR := Y < 0 OR X < 0 OR Y > 23 OR X > 79;

END_FUNCTION

FUNCTION_BLOCK TN_SC_WRITE_ATTR_Block

	VAR
		in_Offset :	INT;
	END_VAR

	VAR_INPUT
		Iin_Y :	INT;
		Iin_X :	INT;
		Iby_ATTR :	BYTE;
	END_VAR

	VAR_IN_OUT
		Xus_TN_SCREEN :	us_TN_SCREEN;
	END_VAR

	IF TN_SC_XY_ERROR(Iin_X,Iin_Y) THEN RETURN; END_IF;
	in_Offset := (Iin_Y * 80) + Iin_X;
	Xus_TN_SCREEN.bya_COLOR[in_Offset] := Iby_ATTR;

END_FUNCTION_BLOCK

PROGRAM program0
	VAR
		Iin_Y :	INT;
		Iin_X :	INT;
		Iby_ATTR :	BYTE;
		Xus_TN_SCREEN :	us_TN_SCREEN;

		func_block : TN_SC_WRITE_ATTR_Block;
	END_VAR
	func_block.Iin_Y := Iin_Y;
	func_block.Iin_X := Iin_X;
	func_block.Iby_ATTR := Iby_ATTR;
	func_block.Xus_TN_SCREEN := Xus_TN_SCREEN;

	func_block();
	Xus_TN_SCREEN  := func_block.Xus_TN_SCREEN;
END_PROGRAM

CONFIGURATION Config0
	RESOURCE Res0 ON PLC
		TASK task0(INTERVAL := T#20ms,PRIORITY := 0);
		PROGRAM instance0 WITH task0 : program0;
	END_RESOURCE
END_CONFIGURATION

(* ---- TN_SC_WRITE_C.ST ---- *)
TYPE
  bya_TN_CHAR:       	ARRAY [0..1919] OF BYTE;
  bya_TN_BACKUP:     	ARRAY [0..1919] OF BYTE;
  bya_TN_COLOR:      	ARRAY [0..1919] OF BYTE;
  bya_TN_Line_Update:	ARRAY [0..23]   OF BOOL;

  us_TN_SCREEN :
  STRUCT
		bya_CHAR:			bya_TN_CHAR;
		bya_COLOR:			bya_TN_COLOR;
		bya_BACKUP:			bya_TN_BACKUP;
		bya_Line_Update:	bya_TN_Line_Update;

		by_Input_Exten_Code:    BYTE;
		by_Input_ASCII_Code:    BYTE;
		bo_Input_ASCII_IsNum:   BOOL;
		in_Page_Number:        	INT;                (* aktive Seiten-Nr.              *)
		in_Cursor_X:           	INT;                (* Cursor X-Position              *)
		in_Cursor_Y:           	INT;                (* Cursor Y-Position              *)
		in_EOS_Offset:         	INT;                (* End of String Offset           *)
		by_Clear_Screen_Attr:  	BYTE;               (* Clear-Screen Attr              *)
		bo_Clear_Screen:       	BOOL;               (* Clear-Screen ausl�sen          *)
		bo_Modal_Dialog:       	BOOL;               (* Modaler Dialog ist aktiv       *)
		bo_Menue_Bar_Dialog:   	BOOL;               (* Menue Dialog ist aktiv         *)

  END_STRUCT;
END_TYPE

FUNCTION _BYTE_TO_INT:INT
	VAR_INPUT
		IN :	BYTE;
	END_VAR

	_BYTE_TO_INT := USINT_TO_INT(BYTE_TO_USINT(IN));
END_FUNCTION

FUNCTION_BLOCK CHR_TO_STRING_Block
	VAR_INPUT
		C :	BYTE;
	END_VAR

	VAR_OUTPUT
		CHR_TO_STRING :	STRING;
	END_VAR

	CHR_TO_STRING := BYTE_TO_STRING(C);

END_FUNCTION_BLOCK

FUNCTION BIT_OF_DWORD : BOOL
  VAR_INPUT
    IN : DWORD;
    N : INT;
  END_VAR

  BIT_OF_DWORD := (SHR(in,N) AND 16#00000001) > 0;
  (* from OSCAT library; www.oscat.de  *)
END_FUNCTION

FUNCTION_BLOCK FILL_Block
	VAR_INPUT
		C :	BYTE;
		L :	INT;
	END_VAR

	VAR_OUTPUT
		FILL :	STRING;
	END_VAR

	VAR
		N :	BYTE;
		I :	INT;
		sx :	STRING;
		CHR_TO_STRING :	CHR_TO_STRING_Block;
		FILL_tmp :	STRING;
	END_VAR

	CHR_TO_STRING(C:=c);
	Sx:=CHR_TO_STRING.CHR_TO_STRING;
	(* create string *)
	N := INT_TO_BYTE(LIMIT(0,L,80));
	(* create a string of characters to be connected to str *)
	FILL := '';
	FOR i := 1 TO 8 DO
		FILL_tmp := FILL;
		FILL := CONCAT(FILL_tmp,FILL);
		IF BIT_OF_DWORD(BYTE_TO_DWORD(N),7) THEN FILL := CONCAT(FILL,Sx); END_IF;
		N := SHL(N,1);
	END_FOR;
END_FUNCTION_BLOCK

FUNCTION_BLOCK FIX_Block

	VAR_INPUT
		STR :	STRING;
		L :	INT;
		C :	BYTE;
		M :	INT;
	END_VAR

	VAR_OUTPUT
		FIX :	STRING;
	END_VAR

	VAR
		N :	INT;
		FILL :	FILL_Block;
	END_VAR

	N := LIMIT(0,L,255) - LEN(str);
	IF N <= 0 THEN
		(* truncate the string at length N *)
		IF M = 1 THEN
			FIX := RIGHT(str,L);
		ELSE
			FIX := LEFT(str,L);
		END_IF;
	ELSIF M = 1 THEN
		(* connect fill characters at the beginning *)
		FILL(C:=C,L:=N);
		FIX := CONCAT(FILL.FILL,str);
	ELSIF M = 2 THEN
		(* center str beween fill characters *)
		(* for an uneven number of fill characters, there is one more at the end *)
		FILL(C:=C,L:=_BYTE_TO_INT(SHR(INT_TO_BYTE(N+1),1)));
		FIX := CONCAT(str,FILL.FILL);
		FILL(C:=C,L:=_BYTE_TO_INT(SHR(INT_TO_BYTE(N),1)));
		FIX := CONCAT(FILL.FILL,FIX);
	ELSE
		(* connect fill characters at the end *)
		FILL(C:=C,L:=N);
		FIX := CONCAT(str,FILL.FILL);
	END_IF;

END_FUNCTION_BLOCK

FUNCTION_BLOCK TN_SC_WRITE_C_Block

	VAR
		FB_FIX :	FIX_Block;
		FB_TN_SC_WRITE :	TN_SC_WRITE;
	END_VAR

	VAR_INPUT
		Iin_Y :	INT;
		Iin_X :	INT;
		Iby_ATTR :	BYTE;
		Ist_STRING :	STRING;
		Iin_LENGTH :	INT;
		Iin_OPTION :	INT;
	END_VAR

	VAR_IN_OUT
		Xus_TN_SCREEN :	us_TN_SCREEN;
	END_VAR

	FB_FIX.str:=Ist_STRING;
	FB_FIX.L:=Iin_LENGTH;
	FB_FIX.C:=BYTE#32;
	FB_FIX.M:=Iin_OPTION;
	FB_FIX();

	FB_TN_SC_WRITE.Iin_Y			:= Iin_Y;
	FB_TN_SC_WRITE.Iin_X			:= Iin_X;
	FB_TN_SC_WRITE.Iby_ATTR			:= Iby_ATTR;
	FB_TN_SC_WRITE.Ist_STRING		:= FB_FIX.FIX;
	FB_TN_SC_WRITE.Xus_TN_SCREEN	:= Xus_TN_SCREEN;
	FB_TN_SC_WRITE();
	Xus_TN_SCREEN := FB_TN_SC_WRITE.Xus_TN_SCREEN;

END_FUNCTION_BLOCK

PROGRAM program0
	VAR
		Iin_Y :	INT;
		Iin_X :	INT;
		Iby_CHAR :	BYTE;
		Xus_TN_SCREEN :	us_TN_SCREEN;

		func_block : TN_SC_WRITE_C_Block;
	END_VAR
	func_block.Iin_Y := Iin_Y;
	func_block.Iin_X := Iin_X;
	func_block.Iby_CHAR := Iby_CHAR;
	func_block.Xus_TN_SCREEN := Xus_TN_SCREEN;

	func_block();
	Xus_TN_SCREEN  := func_block.Xus_TN_SCREEN;
END_PROGRAM

CONFIGURATION Config0
	RESOURCE Res0 ON PLC
		TASK task0(INTERVAL := T#20ms,PRIORITY := 0);
		PROGRAM instance0 WITH task0 : program0;
	END_RESOURCE
END_CONFIGURATION

(* ---- TN_SC_WRITE_CHAR.ST ---- *)
TYPE
  bya_TN_CHAR:       	ARRAY [0..1919] OF BYTE;
  bya_TN_BACKUP:     	ARRAY [0..1919] OF BYTE;
  bya_TN_COLOR:      	ARRAY [0..1919] OF BYTE;
  bya_TN_Line_Update:	ARRAY [0..23]   OF BOOL;

  us_TN_SCREEN :
  STRUCT
		bya_CHAR:			bya_TN_CHAR;
		bya_COLOR:			bya_TN_COLOR;
		bya_BACKUP:			bya_TN_BACKUP;
		bya_Line_Update:	bya_TN_Line_Update;

		by_Input_Exten_Code:    BYTE;
		by_Input_ASCII_Code:    BYTE;
		bo_Input_ASCII_IsNum:   BOOL;
		in_Page_Number:        	INT;                (* aktive Seiten-Nr.              *)
		in_Cursor_X:           	INT;                (* Cursor X-Position              *)
		in_Cursor_Y:           	INT;                (* Cursor Y-Position              *)
		in_EOS_Offset:         	INT;                (* End of String Offset           *)
		by_Clear_Screen_Attr:  	BYTE;               (* Clear-Screen Attr              *)
		bo_Clear_Screen:       	BOOL;               (* Clear-Screen ausl�sen          *)
		bo_Modal_Dialog:       	BOOL;               (* Modaler Dialog ist aktiv       *)
		bo_Menue_Bar_Dialog:   	BOOL;               (* Menue Dialog ist aktiv         *)

  END_STRUCT;
END_TYPE

FUNCTION TN_SC_XY_ERROR:BOOL

	VAR_INPUT
		X :	INT;
		Y :	INT;
	END_VAR

	TN_SC_XY_ERROR := Y < 0 OR X < 0 OR Y > 23 OR X > 79;

END_FUNCTION

FUNCTION_BLOCK TN_SC_WRITE_CHAR_Block

	VAR
		in_Offset :	INT;
	END_VAR

	VAR_INPUT
		Iin_Y :	INT;
		Iin_X :	INT;
		Iby_CHAR :	BYTE;
	END_VAR

	VAR_IN_OUT
		Xus_TN_SCREEN :	us_TN_SCREEN;
	END_VAR

	IF TN_SC_XY_ERROR(Iin_X,Iin_Y) THEN RETURN; END_IF;
	in_Offset := (Iin_Y * 80) + Iin_X;
	Xus_TN_SCREEN.bya_CHAR[in_Offset] := Iby_CHAR;

END_FUNCTION_BLOCK

PROGRAM program0
	VAR
		Iin_Y :	INT;
		Iin_X :	INT;
		Iby_CHAR :	BYTE;
		Xus_TN_SCREEN :	us_TN_SCREEN;

		func_block : TN_SC_WRITE_CHAR_Block;
	END_VAR
	func_block.Iin_Y := Iin_Y;
	func_block.Iin_X := Iin_X;
	func_block.Iby_CHAR := Iby_CHAR;
	func_block.Xus_TN_SCREEN := Xus_TN_SCREEN;

	func_block();
	Xus_TN_SCREEN  := func_block.Xus_TN_SCREEN;
END_PROGRAM

CONFIGURATION Config0
	RESOURCE Res0 ON PLC
		TASK task0(INTERVAL := T#20ms,PRIORITY := 0);
		PROGRAM instance0 WITH task0 : program0;
	END_RESOURCE
END_CONFIGURATION

(* ---- TN_SC_WRITE_EOS.ST ---- *)
TYPE
  bya_TN_CHAR:       	ARRAY [0..1919] OF BYTE;
  bya_TN_BACKUP:     	ARRAY [0..1919] OF BYTE;
  bya_TN_COLOR:      	ARRAY [0..1919] OF BYTE;
  bya_TN_Line_Update:	ARRAY [0..23]   OF BOOL;

  us_TN_SCREEN :
  STRUCT
		bya_CHAR:			bya_TN_CHAR;
		bya_COLOR:			bya_TN_COLOR;
		bya_BACKUP:			bya_TN_BACKUP;
		bya_Line_Update:	bya_TN_Line_Update;

		by_Input_Exten_Code:    BYTE;
		by_Input_ASCII_Code:    BYTE;
		bo_Input_ASCII_IsNum:   BOOL;
		in_Page_Number:        	INT;                (* aktive Seiten-Nr.              *)
		in_Cursor_X:           	INT;                (* Cursor X-Position              *)
		in_Cursor_Y:           	INT;                (* Cursor Y-Position              *)
		in_EOS_Offset:         	INT;                (* End of String Offset           *)
		by_Clear_Screen_Attr:  	BYTE;               (* Clear-Screen Attr              *)
		bo_Clear_Screen:       	BOOL;               (* Clear-Screen ausl�sen          *)
		bo_Modal_Dialog:       	BOOL;               (* Modaler Dialog ist aktiv       *)
		bo_Menue_Bar_Dialog:   	BOOL;               (* Menue Dialog ist aktiv         *)

  END_STRUCT;
END_TYPE

FUNCTION_BLOCK TN_SC_WRITE_EOS_Block

	VAR
		TN_SC_WRITE :	TN_SC_WRITE;
	END_VAR

	VAR_INPUT
		Iby_ATTR :	BYTE;
		Ist_STRING :	STRING;
	END_VAR

	VAR_IN_OUT
		Xus_TN_SCREEN :	us_TN_SCREEN;
	END_VAR

	TN_SC_WRITE.Iin_Y			:= Xus_TN_SCREEN.us_SYS.in_EOS_Offset / 80;
	TN_SC_WRITE.Iin_X			:= Xus_TN_SCREEN.us_SYS.in_EOS_Offset MOD 80;
	TN_SC_WRITE.Iby_ATTR		:= Iby_ATTR;
	TN_SC_WRITE.Ist_STRING		:= Ist_STRING;
	TN_SC_WRITE.Xus_TN_SCREEN	:= Xus_TN_SCREEN;
	TN_SC_WRITE();
	Xus_TN_SCREEN := TN_SC_WRITE.Xus_TN_SCREEN;

END_FUNCTION_BLOCK

PROGRAM program0
	VAR
		Iby_ATTR :	BYTE;
		Ist_STRING :	STRING;

		func_block : TN_SC_WRITE_EOS_Block;
	END_VAR
	func_block.Iby_ATTR := Iby_ATTR;
	func_block.Ist_STRING := Ist_STRING;
	func_block.Xus_TN_SCREEN := Xus_TN_SCREEN;

	func_block();
	URL_TO_STRING  := func_block.URL_TO_STRING;
END_PROGRAM

CONFIGURATION Config0
	RESOURCE Res0 ON PLC
		TASK task0(INTERVAL := T#20ms,PRIORITY := 0);
		PROGRAM instance0 WITH task0 : program0;
	END_RESOURCE
END_CONFIGURATION

(* ---- TN_SEND_ROWS.ST ---- *)
TYPE
  oscat_IP_FIFO128_DATA  : ARRAY [1..128] OF BYTE;
  oscat_Mailbox  : ARRAY [1..16] OF BYTE;

  oscat_IP_FIFO_DATA :
  STRUCT
    X       : oscat_IP_FIFO128_DATA; (* IP_ID FIFO Speicher          *)
    Y       : oscat_IP_FIFO128_DATA; (* IP_ID Z�hler                 *)
    ID      : BYTE;                  (* h�chste vergabene id         *)
    MAX_ID  : BYTE;                  (* maximal Anmeldungen pro ID   *)
    INIT    : BOOL;                  (* Initialisierung durchgef�hrt *)
    EMPTY   : BOOL;                  (* FIFO leer                    *)
    FULL    : BOOL;                  (* FIFO voll                    *)
    TOP     : INT;                   (* maximale anzahl in FIFO      *)
    NW      : INT;                   (* Schreibzeiger                *)
    NR      : INT;                   (* Lesezeiger                   *)
  END_STRUCT;

  oscat_IP_C:
  STRUCT
    C_MODE:			BYTE;          		(*W Mode: TCP/UCP AKTIV/PASSIV                               *)
    C_PORT:         WORD;          		(*W Portnummer                                               *)
    C_IP:           DWORD;         		(*W IP-Adresse gepackt wwxxyyzz = www.xxx.yyy.zzz            *)
    C_STATE:        BYTE;          		(*R Verbindungsstatus ON/OFF + Flanke ON/OFF                 *)
    C_ENABLE:       BOOL;          		(*W Freigabe f�r Connect                                     *)
    R_OBSERVE:      BOOL;          		(*W Empfang ueberwachen                                      *)
    TIME_RESET:     BOOL;          		(*W Alle Timer ruecksetzen                                   *)
    ERROR:          DWORD;         		(*R vvwwxxyy (vv = CON_ERROR, ww = SEN_ERROR, xx = REC_ERROR *)
    FIFO:           oscat_IP_FIFO_DATA; (*I IP FIFO Struktur                                         *)
    MAILBOX:		oscat_Mailbox;		(*I Mailbox: Datenbereich f�r Bausteindatenaustausch         *)
    END_STRUCT;
END_TYPE

TYPE

  oscat_NW_BUF_LONG  : ARRAY [0..4095] OF BYTE;

  oscat_NETWORK_BUFFER :
  STRUCT
    SIZE   : UINT;
    BUFFER : oscat_NW_BUF_LONG;
  END_STRUCT;

END_TYPE

TYPE

  bya_TN_CHAR:       	ARRAY [0..1919] OF BYTE;
  bya_TN_BACKUP:     	ARRAY [0..1919] OF BYTE;
  bya_TN_COLOR:      	ARRAY [0..1919] OF BYTE;
  bya_TN_Line_Update:	ARRAY [0..23]   OF BOOL;

  us_TN_SCREEN :
  STRUCT
    bya_CHAR:			bya_TN_CHAR;
    bya_COLOR:			bya_TN_COLOR;
    bya_BACKUP:			bya_TN_BACKUP;
    bya_Line_Update:	bya_TN_Line_Update;

    by_Input_Exten_Code:    BYTE;
    by_Input_ASCII_Code:    BYTE;
    bo_Input_ASCII_IsNum:   BOOL;
    in_Page_Number:        	INT;                (* aktive Seiten-Nr.              *)
    in_Cursor_X:           	INT;                (* Cursor X-Position              *)
    in_Cursor_Y:           	INT;                (* Cursor Y-Position              *)
    in_EOS_Offset:         	INT;                (* End of String Offset           *)
    by_Clear_Screen_Attr:  	BYTE;               (* Clear-Screen Attr              *)
    bo_Clear_Screen:       	BOOL;               (* Clear-Screen ausl�sen          *)
    bo_Modal_Dialog:       	BOOL;               (* Modaler Dialog ist aktiv       *)
    bo_Menue_Bar_Dialog:   	BOOL;               (* Menue Dialog ist aktiv         *)

  END_STRUCT;
END_TYPE

FUNCTION INT_TO_BCDC:BYTE

	VAR_INPUT
		IN :	INT;
	END_VAR

	INT_TO_BCDC := SHL(INT_TO_BYTE(IN / INT#10),4) OR INT_TO_BYTE(in MOD INT#10);

END_FUNCTION

FUNCTION_BLOCK TN_SEND_ROWS_Block

  VAR_IN_OUT
    IP_C :	oscat_IP_C;
    S_BUF :	oscat_NETWORK_BUFFER;
    Xus_TN_SCREEN :	us_TN_SCREEN;
  END_VAR

  VAR_INPUT
    S_BUF_SIZE :	INT;
  END_VAR

  VAR
    in_Line_Count :	INT;
    in_Col_Count :	INT;
    in_Last_Row_Index :	INT;
    bo_Break_Loop :	BOOL;
    in_Row_Count :	INT;
    in_Offset :	INT;
    in_Write_Index :	INT;
    in_Write_Index_Backup :	INT;
    by_Cur_Color :	BYTE;
    by_last_Color :	BYTE;
    in_Write_Stop :	INT;
  END_VAR

  IF (IP_C.C_STATE < BYTE#127 OR S_BUF.SIZE > UINT#0) THEN
    RETURN;
  END_IF;

  in_Write_Index := UINT_TO_INT(S_BUF.SIZE) - 1;

  in_Write_Index_Backup := in_Write_Index;

  IF (IP_C.C_STATE = BYTE#254) OR (Xus_TN_SCREEN.bo_Clear_Screen) THEN

    Xus_TN_SCREEN.bo_Clear_Screen := FALSE;

    FOR in_Line_Count := INT#00 TO INT#23 DO
      Xus_TN_SCREEN.bya_Line_Update[in_Line_Count] := TRUE;
    END_FOR;

    in_Write_Index := in_Write_Index + INT#1;
    S_BUF.BUFFER[in_Write_Index] := BYTE#16#1B;
    in_Write_Index := in_Write_Index + INT#1;
    S_BUF.BUFFER[in_Write_Index] := BYTE#16#5B;
    in_Write_Index := in_Write_Index + INT#1;
    S_BUF.BUFFER[in_Write_Index] := BYTE#16#30;
    in_Write_Index := in_Write_Index + INT#1;
    S_BUF.BUFFER[in_Write_Index] := BYTE#16#3B;
    in_Write_Index := in_Write_Index + INT#1;
    S_BUF.BUFFER[in_Write_Index] := BYTE#16#33;

    in_Write_Index := in_Write_Index + INT#1;
    S_BUF.BUFFER[in_Write_Index] := (SHR(Xus_TN_SCREEN.by_Clear_Screen_Attr,4) OR BYTE#16#30);

    in_Write_Index := in_Write_Index + INT#1;
    S_BUF.BUFFER[in_Write_Index] := BYTE#16#3B;
    in_Write_Index := in_Write_Index + INT#1;
    S_BUF.BUFFER[in_Write_Index] := BYTE#16#34;

    in_Write_Index := in_Write_Index + INT#1;
    S_BUF.BUFFER[in_Write_Index] := ((Xus_TN_SCREEN.by_Clear_Screen_Attr AND BYTE#16#07) OR BYTE#16#30);

    in_Write_Index := in_Write_Index + INT#1;
    S_BUF.BUFFER[in_Write_Index] := BYTE#16#6D;

    in_Write_Index := in_Write_Index + INT#1;
    S_BUF.BUFFER[in_Write_Index] := BYTE#16#1B;
    in_Write_Index := in_Write_Index + INT#1;
    S_BUF.BUFFER[in_Write_Index] := BYTE#16#5B;
    in_Write_Index := in_Write_Index + INT#1;
    S_BUF.BUFFER[in_Write_Index] := BYTE#16#32;
    in_Write_Index := in_Write_Index + INT#1;
    S_BUF.BUFFER[in_Write_Index] := BYTE#16#4A;

    in_Write_Index := in_Write_Index + INT#1;
    S_BUF.BUFFER[in_Write_Index] := BYTE#16#1B;
    in_Write_Index := in_Write_Index + INT#1;
    S_BUF.BUFFER[in_Write_Index] := BYTE#16#5B;
    in_Write_Index := in_Write_Index + INT#1;
    S_BUF.BUFFER[in_Write_Index] := BYTE#16#3F;
    in_Write_Index := in_Write_Index + INT#1;
    S_BUF.BUFFER[in_Write_Index] := BYTE#16#37;
    in_Write_Index := in_Write_Index + INT#1;
    S_BUF.BUFFER[in_Write_Index] := BYTE#16#6C;

  END_IF;

  in_Last_Row_Index := INT#0;
  bo_Break_Loop := FALSE;
  in_Write_Stop := S_BUF_SIZE-20;

  FOR in_Line_Count := 0 TO 23 DO

    in_Offset := in_Row_Count * INT#80;

    IF (Xus_TN_SCREEN.bya_Line_Update[in_Row_Count] = TRUE) THEN

      in_Write_Index := in_Write_Index + INT#1;
      S_BUF.BUFFER[in_Write_Index] := BYTE#16#1B;
      in_Write_Index := in_Write_Index + INT#1;
      S_BUF.BUFFER[in_Write_Index] := BYTE#16#5B;

      in_Write_Index := in_Write_Index + INT#1;
      S_BUF.BUFFER[in_Write_Index] :=
        SHR(INT_TO_BCDC(in_Row_Count + INT#1),INT#4) OR BYTE#16#30;

      in_Write_Index := in_Write_Index + INT#1;
      S_BUF.BUFFER[in_Write_Index] :=
        (INT_TO_BCDC(in_Row_Count + INT#1) AND BYTE#16#0F) OR BYTE#16#30;

      in_Write_Index := in_Write_Index + INT#1;
      S_BUF.BUFFER[in_Write_Index] := BYTE#16#3B;
      in_Write_Index := in_Write_Index + INT#1;
      S_BUF.BUFFER[in_Write_Index] := BYTE#16#31;
      in_Write_Index := in_Write_Index + INT#1;
      S_BUF.BUFFER[in_Write_Index] := BYTE#16#48;

      FOR in_Col_Count := 0 TO 79 DO

        by_Cur_Color := Xus_TN_SCREEN.bya_COLOR[in_Offset];
        IF (by_Cur_Color <> by_last_Color) OR (in_Col_Count = INT#00) THEN

          in_Write_Index := in_Write_Index + INT#1;
          S_BUF.BUFFER[in_Write_Index] := BYTE#16#1B;

          in_Write_Index := in_Write_Index + INT#1;
          S_BUF.BUFFER[in_Write_Index] := BYTE#16#5B;

          IF  (((by_Cur_Color AND BYTE#2#10001000) XOR (by_last_Color AND BYTE#2#10001000)) <> BYTE#00) OR (in_Col_Count = 0) THEN

            in_Write_Index := in_Write_Index + INT#1;
            S_BUF.BUFFER[in_Write_Index] := BYTE#16#30;
            in_Write_Index := in_Write_Index + INT#1;
            S_BUF.BUFFER[in_Write_Index] := BYTE#16#3B;

            IF (by_Cur_Color AND BYTE#2#00001000) = BYTE#2#00000000 THEN

              in_Write_Index := in_Write_Index + INT#1;
              S_BUF.BUFFER[in_Write_Index] := BYTE#16#31;
              in_Write_Index := in_Write_Index + INT#1;
              S_BUF.BUFFER[in_Write_Index] := BYTE#16#3B;

            END_IF;

            IF (by_Cur_Color AND BYTE#2#10000000) = BYTE#2#10000000 THEN

              in_Write_Index := in_Write_Index + INT#1;
              S_BUF.BUFFER[in_Write_Index] := BYTE#16#35;
              in_Write_Index := in_Write_Index + INT#1;
              S_BUF.BUFFER[in_Write_Index] := BYTE#16#3B;

            END_IF;

          END_IF;

          in_Write_Index := in_Write_Index + INT#1;
          S_BUF.BUFFER[in_Write_Index] := BYTE#16#33;

          in_Write_Index := in_Write_Index + INT#1;
          S_BUF.BUFFER[in_Write_Index] := ((SHR(by_Cur_Color,4) AND BYTE#2#00000111) OR BYTE#16#30);

          in_Write_Index := in_Write_Index + INT#1;
          S_BUF.BUFFER[in_Write_Index] := BYTE#16#3B;

          in_Write_Index := in_Write_Index + INT#1;
          S_BUF.BUFFER[in_Write_Index] := BYTE#16#34;

          in_Write_Index := in_Write_Index + INT#1;
          S_BUF.BUFFER[in_Write_Index] := ((by_Cur_Color AND BYTE#2#00000111) OR BYTE#16#30);

          in_Write_Index := in_Write_Index + INT#1;
          S_BUF.BUFFER[in_Write_Index] := BYTE#16#6D;

          by_last_Color := by_Cur_Color;

        END_IF;

        IF (in_Write_Index > in_Write_Stop) THEN

          bo_Break_Loop := TRUE;
          EXIT;

        END_IF;

        in_Write_Index := in_Write_Index + INT#1;
        S_BUF.BUFFER[in_Write_Index] := Xus_TN_SCREEN.bya_CHAR[in_Offset];

        in_Offset := in_Offset + INT#01;
      END_FOR;

      IF (bo_Break_Loop = TRUE) THEN

        in_Write_Index := in_Last_Row_Index;

        EXIT;
      END_IF;

      in_Last_Row_Index := in_Write_Index;
      Xus_TN_SCREEN.bya_Line_Update[in_Row_Count] := FALSE;

    END_IF;

    in_Row_Count := in_Row_Count + INT#01;

    IF (in_Row_Count > INT#23) THEN
      in_Row_Count := INT#00;
    END_IF;

  END_FOR;

  IF (bo_Break_Loop = FALSE) THEN

    in_Row_Count := INT#00;

  END_IF;

  IF (in_Write_Index <> in_Write_Index_Backup) THEN

    in_Write_Index := in_Write_Index + INT#1;
    S_BUF.BUFFER[in_Write_Index] := BYTE#16#1B;
    in_Write_Index := in_Write_Index + INT#1;
    S_BUF.BUFFER[in_Write_Index] := BYTE#16#5B;

    in_Write_Index := in_Write_Index + INT#1;
    S_BUF.BUFFER[in_Write_Index] := SHR(INT_TO_BCDC(Xus_TN_SCREEN.in_Cursor_Y + 1),INT#4) OR BYTE#16#30;

    in_Write_Index := in_Write_Index + INT#1;
    S_BUF.BUFFER[in_Write_Index] := (INT_TO_BCDC(Xus_TN_SCREEN.in_Cursor_Y + 1) AND BYTE#16#0F) OR BYTE#16#30;

    in_Write_Index := in_Write_Index + INT#1;
    S_BUF.BUFFER[in_Write_Index] := BYTE#16#3B;

    in_Write_Index := in_Write_Index + INT#1;
    S_BUF.BUFFER[in_Write_Index] := SHR(INT_TO_BCDC(Xus_TN_SCREEN.in_Cursor_X + 1),INT#4) OR BYTE#16#30;

    in_Write_Index := in_Write_Index + INT#1;
    S_BUF.BUFFER[in_Write_Index] := (INT_TO_BCDC(Xus_TN_SCREEN.in_Cursor_X + 1) AND BYTE#16#0F) OR BYTE#16#30;

    in_Write_Index := in_Write_Index + INT#1;
    S_BUF.BUFFER[in_Write_Index] := BYTE#16#48;

  END_IF;

  S_BUF.SIZE := INT_TO_UINT(in_Write_Index + 1);

END_FUNCTION_BLOCK

PROGRAM program0
	VAR
		IP_C :	oscat_IP_C;
    S_BUF :	oscat_NETWORK_BUFFER;
    Xus_TN_SCREEN :	us_TN_SCREEN;
    S_BUF_SIZE :	INT;

		func_block : TN_SEND_ROWS_Block;
	END_VAR
	func_block.IP_C := IP_C;
  func_block.S_BUF := S_BUF;
  func_block.Xus_TN_SCREEN := Xus_TN_SCREEN;
  func_block.S_BUF_SIZE := S_BUF_SIZE;

	func_block();
	IP_C  := func_block.IP_C;
  S_BUF  := func_block.S_BUF;
  Xus_TN_SCREEN  := func_block.Xus_TN_SCREEN;
END_PROGRAM

CONFIGURATION Config0
	RESOURCE Res0 ON PLC
		TASK task0(INTERVAL := T#20ms,PRIORITY := 0);
		PROGRAM instance0 WITH task0 : program0;
	END_RESOURCE
END_CONFIGURATION

(* ---- TO_UML.ST ---- *)
FUNCTION _BYTE_TO_INT:INT
	VAR_INPUT
		IN :	BYTE;
	END_VAR

	_BYTE_TO_INT := USINT_TO_INT(BYTE_TO_USINT(IN));
END_FUNCTION

FUNCTION_BLOCK TO_UML_Block

	VAR_INPUT
		IN :	BYTE;
	END_VAR

	VAR_OUTPUT
		TO_UML :	STRING;
	END_VAR

	CASE _BYTE_TO_INT(in) OF
		196:
			TO_UML := 'Ae';
		214:
			TO_UML := 'Oe';
		220:
			TO_UML := 'Ue';
		223:
			TO_UML := 'ss';
		228:
			TO_UML := 'ae';
		246:
			TO_UML := 'oe';
		252:
			TO_UML := 'ue';
	ELSE
		TO_UML := BYTE_TO_STRING(IN);
	END_CASE;

END_FUNCTION_BLOCK

PROGRAM program0
  VAR
	IN :	BYTE;
	TO_UML :	STRING;
	func_block : TO_UML_Block;
  END_VAR
	func_block.IN  := IN;
	func_block();
	TO_UML := func_block.TO_UML;

END_PROGRAM

CONFIGURATION Config0
	RESOURCE Res0 ON PLC
		TASK task0(INTERVAL := T#20ms,PRIORITY := 0);
		PROGRAM instance0 WITH task0 : program0;
	END_RESOURCE
END_CONFIGURATION

(* ---- TOD_TO_STRING.ST ---- *)
FUNCTION HOUR:INT
	VAR_INPUT
		ITOD :	UDINT;
	END_VAR
	hour := UDINT_TO_INT(itod / UDINT#3600000);
END_FUNCTION

FUNCTION MINUTE:INT

	VAR_INPUT
		ITOD :	UDINT;
	END_VAR

	minute := UDINT_TO_INT((itod / UDINT#60000) - ((itod / UDINT#3600000) * UDINT#60));

END_FUNCTION

FUNCTION_BLOCK TOD_TO_STRING_Block
	VAR_INPUT
		ITOD :	UDINT;
	END_VAR

	VAR_OUTPUT
		TOD_STRING :	STRING;
	END_VAR

	VAR
		st_tmp1 :	STRING;
		st_tmp2 :	STRING;
		cur_hours :	INT;
	END_VAR

	cur_hours := hour(ITOD);
	IF cur_hours = 0 THEN
	st_tmp2 := '%01dh';
	ELSE
	st_tmp2 := '%dh';
	END_IF;

	st_tmp1 := CONCAT(INT_TO_STRING(cur_hours),INT_TO_STRING(minute(ITOD)));
	TOD_STRING := CONCAT(st_tmp1,UDINT_TO_STRING(ITOD MOD UDINT#60000 / UDINT#1000));
END_FUNCTION_BLOCK

PROGRAM program0
  VAR
    LocalVar0 : UDINT;
	LocalOUT  : STRING;
	func_block : TOD_TO_STRING_Block;
  END_VAR
	func_block.ITOD  := LocalVar0;
	func_block();
	LocalOUT := func_block.TOD_STRING;
END_PROGRAM

CONFIGURATION Config0
  RESOURCE Res0 ON PLC
    TASK task0(INTERVAL := T#20ms,PRIORITY := 0);
    PROGRAM instance0 WITH task0 : program0;
  END_RESOURCE
END_CONFIGURATION

(* ---- TOF_1.ST ---- *)
FUNCTION UDINT_TO_TIME2:TIME

	VAR_INPUT
		IN :	UDINT;
	END_VAR

	UDINT_TO_TIME2 := DINT_TO_TIME(UDINT_TO_DINT(IN));

END_FUNCTION

FUNCTION_BLOCK T_PLC_MS_block
	VAR_OUTPUT
		T_PLC_MS :	UDINT;
	END_VAR

	VAR_EXTERNAL
		PLC_TICKS_PER_SEC :	INT;
		PLC_SYS_TICK_CNT :	DINT;
	END_VAR

	VAR
		debug :	BOOL;(*Debug-Mode ON / OFF*)
		N :	INT;(*Debug-Faktor*)
		Offset :	UDINT;(*Debug-Offset*)
		temp :	DWORD := DWORD#1;(*Debug-Offset*)
		mode :	BOOL;(*modus*)
		faktor :	UDINT;(*Systemtakt-Faktor*)
		init :	BOOL;
		v_plc_ticks_per_sec :	UDINT;
		base :	UDINT := UDINT#1000;
	END_VAR

	IF init = FALSE THEN
		v_plc_ticks_per_sec := INT_TO_UDINT(PLC_TICKS_PER_SEC);
		IF v_plc_ticks_per_sec = UDINT#1024 THEN
			faktor := UDINT#1;
			mode := FALSE;
		ELSIF v_plc_ticks_per_sec > UDINT#0 THEN
			IF v_plc_ticks_per_sec <= base THEN
				faktor := base / v_plc_ticks_per_sec;
				mode := FALSE;
			ELSE
				faktor := v_plc_ticks_per_sec / base;
				mode := TRUE;
			END_IF;
		ELSE
			faktor := UDINT#1;
		END_IF;
		init := TRUE;
	END_IF;

	IF mode THEN
		T_PLC_MS := DINT_TO_UDINT(PLC_SYS_TICK_CNT) / faktor;
	ELSE
		T_PLC_MS := DINT_TO_UDINT(PLC_SYS_TICK_CNT) * faktor;
	END_IF;

	IF debug THEN
		T_PLC_MS := (DWORD_TO_UDINT(SHL(UDINT_TO_DWORD(T_PLC_MS),N) OR SHL(temp,N)) - UDINT#1) + Offset;
	END_IF;

END_FUNCTION_BLOCK

FUNCTION_BLOCK TOF_1

	VAR_INPUT
		IN :	BOOL;
		PT :	TIME;
		RST :	BOOL;
	END_VAR

	VAR_OUTPUT
		Q :	BOOL;
	END_VAR

	VAR
		start :	TIME;
		tx :	TIME;
		T_PLC_MS :	T_PLC_MS_block;
	END_VAR

	T_PLC_MS();
	tx:= UDINT_TO_TIME(T_PLC_MS.T_PLC_MS);

	IF RST THEN
		Q := FALSE;
	ELSIF IN THEN
		Q := TRUE;
		start := tx;
	ELSIF tx - start >= PT THEN
		Q := FALSE;
	END_IF;

END_FUNCTION_BLOCK

PROGRAM program0
  VAR
	IN :	BOOL;
	PT :	TIME;
	RST :	BOOL;
	Q :	BOOL;
	func_block : TOF_1;
  END_VAR
	func_block.IN  :=IN;
	func_block.PT  :=PT;
	func_block.RST  :=RST;
	func_block();
	Q := func_block.Q;
END_PROGRAM

CONFIGURATION Config0
	VAR_GLOBAL
		PLC_TICKS_PER_SEC :	INT;
		PLC_SYS_TICK_CNT :	DINT;
	END_VAR
	RESOURCE Res0 ON PLC
		TASK task0(INTERVAL := T#20ms,PRIORITY := 0);
		PROGRAM instance0 WITH task0 : program0;
	END_RESOURCE
END_CONFIGURATION

(* ---- TOGGLE.ST ---- *)
FUNCTION_BLOCK TOGGLE

	VAR_INPUT
		CLK :	BOOL;
		RST :	BOOL;
	END_VAR

	VAR_OUTPUT
		Q :	BOOL;
	END_VAR

	VAR
		edge :	BOOL;
	END_VAR

	IF rst THEN
		Q := FALSE;
	ELSIF clk AND NOT edge THEN
		Q := NOT Q;
	END_IF;
	edge := clk;

END_FUNCTION_BLOCK

PROGRAM program0
  VAR
	CLK :	BOOL;
	RST :	BOOL;
	Q :	BOOL;
	func_block : TOGGLE;
  END_VAR
	func_block.CLK  :=CLK;
	func_block.RST  :=RST;
	func_block();
	Q := func_block.Q;

END_PROGRAM

CONFIGURATION Config0
	RESOURCE Res0 ON PLC
		TASK task0(INTERVAL := T#20ms,PRIORITY := 0);
		PROGRAM instance0 WITH task0 : program0;
	END_RESOURCE
END_CONFIGURATION

(* ---- TONOF.ST ---- *)
FUNCTION_BLOCK TONOF

	VAR_INPUT
		IN :	BOOL;
		T_ON :	TIME;
		T_OFF :	TIME;
	END_VAR

	VAR_OUTPUT
		Q :	BOOL;
	END_VAR

	VAR
		X :	TON;
		old :	BOOL;
		mode :	BOOL;
	END_VAR

	IF IN XOR old THEN
	X(IN := FALSE, PT := SEL_TIME(IN,T_OFF,T_ON));
	mode := IN;
	old := IN;
	END_IF;
	X(IN := TRUE);
	IF X.Q THEN Q := mode;END_IF;

END_FUNCTION_BLOCK

PROGRAM program0
  VAR
	IN :	BOOL;
	T_ON :	TIME;
	T_OFF :	TIME;
	Q :	BOOL;
	func_block : TONOF;
  END_VAR
	func_block.IN  :=IN ;
	func_block.T_ON  :=T_ON ;
	func_block.T_OFF  :=T_OFF ;
	func_block();
	Q := func_block.Q;

END_PROGRAM

CONFIGURATION Config0
	RESOURCE Res0 ON PLC
		TASK task0(INTERVAL := T#20ms,PRIORITY := 0);
		PROGRAM instance0 WITH task0 : program0;
	END_RESOURCE
END_CONFIGURATION

(* ---- TP_1.ST ---- *)
FUNCTION UDINT_TO_TIME2:TIME

	VAR_INPUT
		IN :	UDINT;
	END_VAR

	UDINT_TO_TIME2 := DINT_TO_TIME(UDINT_TO_DINT(IN));

END_FUNCTION

FUNCTION_BLOCK T_PLC_MS_block
	VAR_OUTPUT
		T_PLC_MS :	UDINT;
	END_VAR

	VAR_EXTERNAL
		PLC_TICKS_PER_SEC :	INT;
		PLC_SYS_TICK_CNT :	DINT;
	END_VAR

	VAR
		debug :	BOOL;(*Debug-Mode ON / OFF*)
		N :	INT;(*Debug-Faktor*)
		Offset :	UDINT;(*Debug-Offset*)
		temp :	DWORD := DWORD#1;(*Debug-Offset*)
		mode :	BOOL;(*modus*)
		faktor :	UDINT;(*Systemtakt-Faktor*)
		init :	BOOL;
		v_plc_ticks_per_sec :	UDINT;
		base :	UDINT := UDINT#1000;
	END_VAR

	IF init = FALSE THEN
		v_plc_ticks_per_sec := INT_TO_UDINT(PLC_TICKS_PER_SEC);
		IF v_plc_ticks_per_sec = UDINT#1024 THEN
			faktor := UDINT#1;
			mode := FALSE;
		ELSIF v_plc_ticks_per_sec > UDINT#0 THEN
			IF v_plc_ticks_per_sec <= base THEN
				faktor := base / v_plc_ticks_per_sec;
				mode := FALSE;
			ELSE
				faktor := v_plc_ticks_per_sec / base;
				mode := TRUE;
			END_IF;
		ELSE
			faktor := UDINT#1;
		END_IF;
		init := TRUE;
	END_IF;

	IF mode THEN
		T_PLC_MS := DINT_TO_UDINT(PLC_SYS_TICK_CNT) / faktor;
	ELSE
		T_PLC_MS := DINT_TO_UDINT(PLC_SYS_TICK_CNT) * faktor;
	END_IF;

	IF debug THEN
		T_PLC_MS := (DWORD_TO_UDINT(SHL(UDINT_TO_DWORD(T_PLC_MS),N) OR SHL(temp,N)) - UDINT#1) + Offset;
	END_IF;

END_FUNCTION_BLOCK

FUNCTION_BLOCK TP_1

	VAR_INPUT
		IN :	BOOL;
		PT :	TIME;
		RST :	BOOL;
	END_VAR

	VAR_OUTPUT
		Q :	BOOL;
	END_VAR

	VAR
		tx :	TIME;
		start :	TIME;
		ix :	BOOL;
		T_PLC_MS :	T_PLC_MS_block;
	END_VAR

	T_PLC_MS();
	tx := UDINT_TO_TIME(T_PLC_MS.T_PLC_MS);

	IF RST THEN
		Q := FALSE;
	ELSIF IN AND NOT ix THEN
		Q := TRUE;
		start := tx;
	ELSIF tx - start >= PT THEN
		Q := FALSE;
	END_IF;

	ix:= IN;

END_FUNCTION_BLOCK

PROGRAM program0
  VAR
	IN :	BOOL;
	PT :	TIME;
	RST :	BOOL;
	Q :	BOOL;
	func_block : TP_1;
  END_VAR
	func_block.IN  :=IN;
	func_block.PT  :=PT;
	func_block.RST  :=RST;
	func_block();
	Q := func_block.Q;
END_PROGRAM

CONFIGURATION Config0
	VAR_GLOBAL
		PLC_TICKS_PER_SEC :	INT;
		PLC_SYS_TICK_CNT :	DINT;
	END_VAR
	RESOURCE Res0 ON PLC
		TASK task0(INTERVAL := T#20ms,PRIORITY := 0);
		PROGRAM instance0 WITH task0 : program0;
	END_RESOURCE
END_CONFIGURATION

(* ---- TP_1D.ST ---- *)
FUNCTION UDINT_TO_TIME2:TIME

	VAR_INPUT
		IN :	UDINT;
	END_VAR

	UDINT_TO_TIME2 := DINT_TO_TIME(UDINT_TO_DINT(IN));

END_FUNCTION

FUNCTION_BLOCK T_PLC_MS_block
	VAR_OUTPUT
		T_PLC_MS :	UDINT;
	END_VAR

	VAR_EXTERNAL
		PLC_TICKS_PER_SEC :	INT;
		PLC_SYS_TICK_CNT :	DINT;
	END_VAR

	VAR
		debug :	BOOL;(*Debug-Mode ON / OFF*)
		N :	INT;(*Debug-Faktor*)
		Offset :	UDINT;(*Debug-Offset*)
		temp :	DWORD := DWORD#1;(*Debug-Offset*)
		mode :	BOOL;(*modus*)
		faktor :	UDINT;(*Systemtakt-Faktor*)
		init :	BOOL;
		v_plc_ticks_per_sec :	UDINT;
		base :	UDINT := UDINT#1000;
	END_VAR

	IF init = FALSE THEN
		v_plc_ticks_per_sec := INT_TO_UDINT(PLC_TICKS_PER_SEC);
		IF v_plc_ticks_per_sec = UDINT#1024 THEN
			faktor := UDINT#1;
			mode := FALSE;
		ELSIF v_plc_ticks_per_sec > UDINT#0 THEN
			IF v_plc_ticks_per_sec <= base THEN
				faktor := base / v_plc_ticks_per_sec;
				mode := FALSE;
			ELSE
				faktor := v_plc_ticks_per_sec / base;
				mode := TRUE;
			END_IF;
		ELSE
			faktor := UDINT#1;
		END_IF;
		init := TRUE;
	END_IF;

	IF mode THEN
		T_PLC_MS := DINT_TO_UDINT(PLC_SYS_TICK_CNT) / faktor;
	ELSE
		T_PLC_MS := DINT_TO_UDINT(PLC_SYS_TICK_CNT) * faktor;
	END_IF;

	IF debug THEN
		T_PLC_MS := (DWORD_TO_UDINT(SHL(UDINT_TO_DWORD(T_PLC_MS),N) OR SHL(temp,N)) - UDINT#1) + Offset;
	END_IF;

END_FUNCTION_BLOCK

FUNCTION_BLOCK TP_1D
	VAR_INPUT
		IN :	BOOL;
		PT1 :	TIME;
		PTD :	TIME;
		RST :	BOOL;
	END_VAR

	VAR_OUTPUT
		Q :	BOOL;
		W :	BOOL;
	END_VAR

	VAR
		tx :	TIME;
		start :	TIME;
		ix :	BOOL;
		T_PLC_MS :	T_PLC_MS_block;
	END_VAR

	T_PLC_MS();
	tx := UDINT_TO_TIME(T_PLC_MS.T_PLC_MS);

	IF RST THEN
		Q := FALSE;
		rst := FALSE;
		W := FALSE;
	ELSIF W THEN
		IF tx - start >= PTD THEN
			W := FALSE;
		END_IF;
	ELSIF IN AND NOT ix THEN
		Q := TRUE;
		start := tx;
		in := FALSE;
	ELSIF tx - start >= PT1 THEN
		Q := FALSE;
		W := TRUE;
		start := tx;
	END_IF;

	ix := IN;

END_FUNCTION_BLOCK

PROGRAM program0
  VAR
	IN :	BOOL;
	PT1 :	TIME;
	PTD :	TIME;
	RST :	BOOL;
	Q :	BOOL;
	W :	BOOL;
	func_block : TP_1D;
  END_VAR
	func_block.IN  :=IN;
	func_block.PT1  :=PT1;
	func_block.PTD  :=PTD;
	func_block.RST  :=RST;
	func_block();
	Q := func_block.Q;
	W := func_block.W;
END_PROGRAM

CONFIGURATION Config0
	VAR_GLOBAL
		PLC_TICKS_PER_SEC :	INT;
		PLC_SYS_TICK_CNT :	DINT;
	END_VAR
	RESOURCE Res0 ON PLC
		TASK task0(INTERVAL := T#20ms,PRIORITY := 0);
		PROGRAM instance0 WITH task0 : program0;
	END_RESOURCE
END_CONFIGURATION

(* ---- TP_X.ST ---- *)
FUNCTION UDINT_TO_TIME2:TIME

	VAR_INPUT
		IN :	UDINT;
	END_VAR

	UDINT_TO_TIME2 := DINT_TO_TIME(UDINT_TO_DINT(IN));

END_FUNCTION

FUNCTION_BLOCK T_PLC_MS_block
	VAR_OUTPUT
		T_PLC_MS :	UDINT;
	END_VAR

	VAR_EXTERNAL
		PLC_TICKS_PER_SEC :	INT;
		PLC_SYS_TICK_CNT :	DINT;
	END_VAR

	VAR
		debug :	BOOL;(*Debug-Mode ON / OFF*)
		N :	INT;(*Debug-Faktor*)
		Offset :	UDINT;(*Debug-Offset*)
		temp :	DWORD := DWORD#1;(*Debug-Offset*)
		mode :	BOOL;(*modus*)
		faktor :	UDINT;(*Systemtakt-Faktor*)
		init :	BOOL;
		v_plc_ticks_per_sec :	UDINT;
		base :	UDINT := UDINT#1000;
	END_VAR

	IF init = FALSE THEN
		v_plc_ticks_per_sec := INT_TO_UDINT(PLC_TICKS_PER_SEC);
		IF v_plc_ticks_per_sec = UDINT#1024 THEN
			faktor := UDINT#1;
			mode := FALSE;
		ELSIF v_plc_ticks_per_sec > UDINT#0 THEN
			IF v_plc_ticks_per_sec <= base THEN
				faktor := base / v_plc_ticks_per_sec;
				mode := FALSE;
			ELSE
				faktor := v_plc_ticks_per_sec / base;
				mode := TRUE;
			END_IF;
		ELSE
			faktor := UDINT#1;
		END_IF;
		init := TRUE;
	END_IF;

	IF mode THEN
		T_PLC_MS := DINT_TO_UDINT(PLC_SYS_TICK_CNT) / faktor;
	ELSE
		T_PLC_MS := DINT_TO_UDINT(PLC_SYS_TICK_CNT) * faktor;
	END_IF;

	IF debug THEN
		T_PLC_MS := (DWORD_TO_UDINT(SHL(UDINT_TO_DWORD(T_PLC_MS),N) OR SHL(temp,N)) - UDINT#1) + Offset;
	END_IF;

END_FUNCTION_BLOCK

FUNCTION_BLOCK TP_X
	VAR_INPUT
		IN :	BOOL;
		PT :	TIME;
	END_VAR

	VAR_OUTPUT
		Q :	BOOL;
		ET :	TIME;
	END_VAR

	VAR
		edge :	BOOL;
		start :	TIME;
		tx :	TIME;
		T_PLC_MS :	T_PLC_MS_block;
	END_VAR

	T_PLC_MS();
	tx := UDINT_TO_TIME2(T_PLC_MS.T_PLC_MS);

	IF IN AND NOT edge THEN
		start := tx;
		Q := PT > t#0ms;
	ELSIF Q THEN
		ET := tx - start;
		IF ET >= PT THEN
			Q := FALSE;
			ET := t#0ms;
		END_IF;
	END_IF;
	edge := IN;

END_FUNCTION_BLOCK

PROGRAM program0
  VAR
	IN :	BOOL;
	PT :	TIME;
	Q :	BOOL;
	ET :	TIME;
	func_block : TP_X;
  END_VAR
	func_block.IN  :=IN;
	func_block.PT  :=PT ;
	func_block();
	Q := func_block.Q;
	ET := func_block.ET;
END_PROGRAM

CONFIGURATION Config0
	VAR_GLOBAL
		PLC_TICKS_PER_SEC :	INT;
		PLC_SYS_TICK_CNT :	DINT;
	END_VAR
	RESOURCE Res0 ON PLC
		TASK task0(INTERVAL := T#20ms,PRIORITY := 0);
		PROGRAM instance0 WITH task0 : program0;
	END_RESOURCE
END_CONFIGURATION

(* ---- TREND.ST ---- *)
FUNCTION_BLOCK TREND

	VAR_INPUT
		X :	REAL;
	END_VAR

	VAR_OUTPUT
		Q :	BOOL;
		TU :	BOOL;
		TD :	BOOL;
		D :	REAL;
	END_VAR

	VAR
		last_x :	REAL;
	END_VAR

	TU := X > last_X;
	TD := X < last_X;
	Q := TU OR TD;
	D := X - LAST_X;

	last_X := X;

END_FUNCTION_BLOCK

PROGRAM program0
  VAR
	X :	REAL;
	Q :	BOOL;
	TU :	BOOL;
	TD :	BOOL;
	D :	REAL;
	func_block : TREND;
  END_VAR
	func_block.X  :=X ;
	func_block();
	Q := func_block.Q;
	TU := func_block.TU;
	TD := func_block.TD;
	D := func_block.D;
END_PROGRAM

CONFIGURATION Config0
	RESOURCE Res0 ON PLC
		TASK task0(INTERVAL := T#20ms,PRIORITY := 0);
		PROGRAM instance0 WITH task0 : program0;
	END_RESOURCE
END_CONFIGURATION

(* ---- TREND_DW.ST ---- *)
FUNCTION_BLOCK TREND_DW
	VAR_INPUT
		X :	DWORD;
	END_VAR
	VAR_OUTPUT
		Q :	BOOL;
		TU :	BOOL;
		TD :	BOOL;
		D :	DWORD;
	END_VAR

	VAR
		LAST_X :	DWORD;
	END_VAR

	IF X > last_X THEN
		TU := TRUE;
		TD := FALSE;
		D := UDINT_TO_DWORD(DWORD_TO_UDINT(X) - DWORD_TO_UDINT(last_X));
		Q := TRUE;
	ELSIF X < last_X THEN
		TD := TRUE;
		TU := FALSE;
		D := UDINT_TO_DWORD(DWORD_TO_UDINT(last_X) - DWORD_TO_UDINT(X));
		Q := FALSE;
	ELSE
		TU := FALSE;
		TD := FALSE;
		D := DWORD#0;
	END_IF;
	last_X := X;
END_FUNCTION_BLOCK

PROGRAM program0
  VAR
	X :	DWORD;
	Q :	BOOL;
	TU :	BOOL;
	TD :	BOOL;
	D :	DWORD;
	func_block : TREND_DW;
  END_VAR
	func_block.X  :=X ;
	func_block();
	Q := func_block.Q;
	TU := func_block.TU;
	TD := func_block.TD;
	D := func_block.D;
END_PROGRAM

CONFIGURATION Config0
	RESOURCE Res0 ON PLC
		TASK task0(INTERVAL := T#20ms,PRIORITY := 0);
		PROGRAM instance0 WITH task0 : program0;
	END_RESOURCE
END_CONFIGURATION

(* ---- TRIM.ST ---- *)
FUNCTION_BLOCK TRIM

	VAR_INPUT
		STR :	STRING;
	END_VAR

	VAR_OUTPUT
		TRIM3 :	STRING;
	END_VAR

	VAR
		pos :	INT;
	END_VAR

	trim3 := str;
	REPEAT
		pos := FIND(trim3,' ');
		IF pos > 0 THEN trim3 := REPLACE(trim3,'',1,pos); END_IF;
	UNTIL pos = 0 END_REPEAT;

END_FUNCTION_BLOCK

PROGRAM program0
  VAR
	STR :	STRING;

	TRIM3 :	STRING;
	func_block : TRIM;
  END_VAR
	func_block.STR  :=STR ;
	func_block();
	TRIM3 := func_block.TRIM3;

END_PROGRAM

CONFIGURATION Config0
	RESOURCE Res0 ON PLC
		TASK task0(INTERVAL := T#20ms,PRIORITY := 0);
		PROGRAM instance0 WITH task0 : program0;
	END_RESOURCE
END_CONFIGURATION

(* ---- TRIM1.ST ---- *)
FUNCTION_BLOCK TRIM1

	VAR_INPUT
		STR :	STRING;
	END_VAR

	VAR_OUTPUT
		TRIM3 :	STRING;
	END_VAR

	VAR
		pos :	INT;
		st_temp :	STRING;
	END_VAR

	trim3 := str;
	REPEAT
		pos := FIND(trim3,'  ');
		IF pos > 0 THEN
		st_temp := trim3;
		trim3 := REPLACE(trim3,' ',2,pos);
		END_IF;
	UNTIL pos = 0 END_REPEAT;
	st_temp := LEFT(trim3,1);
	IF EQ_STRING(st_temp,' ') THEN trim3 := DELETE(trim3,1,1); END_IF;
	st_temp := RIGHT(trim3,1);
	IF EQ_STRING(st_temp,' ') THEN trim3 := DELETE(trim3,1,LEN(trim3)); END_IF;

END_FUNCTION_BLOCK

PROGRAM program0
  VAR
	STR :	STRING;

	TRIM3 :	STRING;
	func_block : TRIM1;
  END_VAR
	func_block.STR  :=STR ;
	func_block();
	TRIM3 := func_block.TRIM3;

END_PROGRAM

CONFIGURATION Config0
	RESOURCE Res0 ON PLC
		TASK task0(INTERVAL := T#20ms,PRIORITY := 0);
		PROGRAM instance0 WITH task0 : program0;
	END_RESOURCE
END_CONFIGURATION

(* ---- TRIME.ST ---- *)
FUNCTION_BLOCK TRIME_Block
	VAR_INPUT
		STR :	STRING;
	END_VAR

	VAR_OUTPUT
		TRIME :	STRING;
	END_VAR

	TRIME := str;
	IF LEN(TRIME) < 1 THEN RETURN; END_IF;

	WHILE (GET_CHAR(TRIME,1) = 32) DO
		TRIME := DELETE(TRIME,1,1);
	END_WHILE;

	WHILE (GET_CHAR(TRIME,LEN(TRIME)) = 32) DO
		TRIME := DELETE(TRIME,1,LEN(TRIME));
	END_WHILE;

END_FUNCTION_BLOCK

PROGRAM program0
  	VAR
		INPUT_STR :	STRING;
		OUTPUT_TRIME : STRING;
		func_block : TRIME_Block;
  	END_VAR
	func_block.STR := INPUT_STR;
	func_block();
	OUTPUT_TRIME := func_block.TRIME;
END_PROGRAM

CONFIGURATION Config0
	RESOURCE Res0 ON PLC
		TASK task0(INTERVAL := T#20ms,PRIORITY := 0);
		PROGRAM instance0 WITH task0 : program0;
	END_RESOURCE
END_CONFIGURATION

(* ---- TUNE.ST ---- *)
FUNCTION_BLOCK T_PLC_MS_Block
	VAR_OUTPUT
		T_PLC_MS :	UDINT;
	END_VAR

	VAR_EXTERNAL
		PLC_TICKS_PER_SEC :	INT;
		PLC_SYS_TICK_CNT :	DINT;
	END_VAR

	VAR
		debug :	BOOL;(*Debug-Mode ON / OFF*)
		N :	INT;(*Debug-Faktor*)
		Offset :	UDINT;(*Debug-Offset*)
		temp :	DWORD := DWORD#1;(*Debug-Offset*)
		mode :	BOOL;(*modus*)
		faktor :	UDINT;(*Systemtakt-Faktor*)
		init :	BOOL;
		v_plc_ticks_per_sec :	UDINT;
		base :	UDINT := UDINT#1000;
	END_VAR

	IF init = FALSE THEN
		v_plc_ticks_per_sec := INT_TO_UDINT(PLC_TICKS_PER_SEC);
		IF v_plc_ticks_per_sec = UDINT#1024 THEN
			faktor := UDINT#1;
			mode := FALSE;
		ELSIF v_plc_ticks_per_sec > UDINT#0 THEN
			IF v_plc_ticks_per_sec <= base THEN
				faktor := base / v_plc_ticks_per_sec;
				mode := FALSE;
			ELSE
				faktor := v_plc_ticks_per_sec / base;
				mode := TRUE;
			END_IF;
		ELSE
			faktor := UDINT#1;
		END_IF;
		init := TRUE;
	END_IF;

	IF mode THEN
		T_PLC_MS := DINT_TO_UDINT(PLC_SYS_TICK_CNT) / faktor;
	ELSE
		T_PLC_MS := DINT_TO_UDINT(PLC_SYS_TICK_CNT) * faktor;
	END_IF;

	IF debug THEN
		T_PLC_MS := (DWORD_TO_UDINT(SHL(UDINT_TO_DWORD(T_PLC_MS),N) OR SHL(temp,N)) - UDINT#1) + Offset;
	END_IF;
END_FUNCTION_BLOCK

FUNCTION TIME_TO_UDINT2:UDINT
	VAR_INPUT
		X :	TIME;
	END_VAR

	TIME_TO_UDINT2 := DINT_TO_UDINT(TIME_TO_DINT(X));
END_FUNCTION

FUNCTION_BLOCK TUNE_Block

	VAR_INPUT
		SET :	BOOL;
		SU :	BOOL;
		SD :	BOOL;
		RST :	BOOL;
		SS :	REAL := 0.1;
		LIMIT_L :	REAL;
		LIMIT_H :	REAL := 100.0;
		RST_VAL :	REAL;
		SET_VAL :	REAL := 100.0;
		T1 :	TIME := T#500ms;
		T2 :	TIME := T#2s;
		S1 :	REAL := 2.0;
		S2 :	REAL := 10.0;
	END_VAR

	VAR_OUTPUT
		Y :	REAL;
	END_VAR

	VAR
		tx :	UDINT;
		start :	UDINT;
		start2 :	UDINT;
		state :	INT;
		in :	BOOL;
		step2 :	REAL;
		speed :	REAL;
		Y_start :	REAL;
		Y_start2 :	REAL;
		T_PLC_MS :	T_PLC_MS_Block;
	END_VAR

	T_PLC_MS();
	tx:= T_PLC_MS.T_PLC_MS;

	IF rst THEN
		Y := RST_val;
		state := 0;
	ELSIF set THEN
		Y := SET_val;
		state := 0;
	ELSIF state > 0 THEN
		IF state = 1 THEN
			in := su;
		ELSE
			in := sd;
		END_IF;
		IF NOT in AND tx - start <= TIME_TO_UDINT2(T1) THEN
			Y := Y_start + step2;
			state := 0;
		ELSIF in AND tx - start >= TIME_TO_UDINT2(T2) THEN
			Y := Y_start2 + UDINT_TO_REAL(tx - start2) * s2 / speed;
		ELSIF in AND tx - start >= TIME_TO_UDINT2(T1) THEN
			Y := Y_start + UDINT_TO_REAL(tx - start - TIME_TO_UDINT2(T1)) * S1 / speed;
			start2 := tx;
			Y_start2 := Y;
		ELSIF NOT in THEN
			state := 0;
		END_IF;
	ELSIF su THEN
		state := 1;
		start := tx;
		step2 := ss;
		speed := 1000.0;
		Y_start := Y;
	ELSIF sd THEN

		state := 2;
		start := tx;
		step2 := -ss;
		speed := -1000.0;
		Y_start := Y;
	END_IF;

END_FUNCTION_BLOCK

PROGRAM program0
  	VAR
		SET :	BOOL;
		SU :	BOOL;
		SD :	BOOL;
		RST :	BOOL;
		SS :	REAL := 0.1;
		LIMIT_L :	REAL;
		LIMIT_H :	REAL := 100.0;
		RST_VAL :	REAL;
		SET_VAL :	REAL := 100.0;
		T1 :	TIME := T#500ms;
		T2 :	TIME := T#2s;
		S1 :	REAL := 2.0;
		S2 :	REAL := 10.0;
		Y :	REAL;
		func_block : TUNE_Block;
  	END_VAR
	func_block.SET := SET;
	func_block.SU := SU;
	func_block.SD := SD;
	func_block.RST := RST;
	func_block.SS:= SS;
	func_block.LIMIT_L := LIMIT_L;
	func_block.LIMIT_H := LIMIT_H;
	func_block.RST_VAL := RST_VAL;
	func_block.SET_VAL := SET_VAL;
	func_block.T1 := T1;
	func_block.T2 := T2;
	func_block.S1 := S1;
	func_block.S2 := S2;
	func_block();
	Y := func_block.Y;
END_PROGRAM

CONFIGURATION Config0
	VAR_GLOBAL
		PLC_TICKS_PER_SEC :	INT;
		PLC_SYS_TICK_CNT :	DINT;
	END_VAR
	RESOURCE Res0 ON PLC
		TASK task0(INTERVAL := T#20ms,PRIORITY := 0);
		PROGRAM instance0 WITH task0 : program0;
	END_RESOURCE
END_CONFIGURATION

(* ---- TUNE2.ST ---- *)
FUNCTION_BLOCK T_PLC_MS_block
	VAR_OUTPUT
		T_PLC_MS :	UDINT;
	END_VAR

	VAR_EXTERNAL
		PLC_TICKS_PER_SEC :	INT;
		PLC_SYS_TICK_CNT :	DINT;
	END_VAR

	VAR
		debug :	BOOL;(*Debug-Mode ON / OFF*)
		N :	INT;(*Debug-Faktor*)
		Offset :	UDINT;(*Debug-Offset*)
		temp :	DWORD := DWORD#1;(*Debug-Offset*)
		mode :	BOOL;(*modus*)
		faktor :	UDINT;(*Systemtakt-Faktor*)
		init :	BOOL;
		v_plc_ticks_per_sec :	UDINT;
		base :	UDINT := UDINT#1000;
	END_VAR

	IF init = FALSE THEN
		v_plc_ticks_per_sec := INT_TO_UDINT(PLC_TICKS_PER_SEC);
		IF v_plc_ticks_per_sec = UDINT#1024 THEN
			faktor := UDINT#1;
			mode := FALSE;
		ELSIF v_plc_ticks_per_sec > UDINT#0 THEN
			IF v_plc_ticks_per_sec <= base THEN
				faktor := base / v_plc_ticks_per_sec;
				mode := FALSE;
			ELSE
				faktor := v_plc_ticks_per_sec / base;
				mode := TRUE;
			END_IF;
		ELSE
			faktor := UDINT#1;
		END_IF;
		init := TRUE;
	END_IF;

	IF mode THEN
		T_PLC_MS := DINT_TO_UDINT(PLC_SYS_TICK_CNT) / faktor;
	ELSE
		T_PLC_MS := DINT_TO_UDINT(PLC_SYS_TICK_CNT) * faktor;
	END_IF;

	IF debug THEN
		T_PLC_MS := (DWORD_TO_UDINT(SHL(UDINT_TO_DWORD(T_PLC_MS),N) OR SHL(temp,N)) - UDINT#1) + Offset;
	END_IF;
END_FUNCTION_BLOCK

FUNCTION TIME_TO_UDINT2:UDINT
	VAR_INPUT
		X :	TIME;
	END_VAR

	TIME_TO_UDINT2 := DINT_TO_UDINT(TIME_TO_DINT(X));
END_FUNCTION

FUNCTION_BLOCK TUNE2_Block

	VAR_INPUT
		SET :	BOOL;
		SU :	BOOL;
		SD :	BOOL;
		FU :	BOOL;
		FD :	BOOL;
		RST :	BOOL;
		SS :	REAL := 0.1;
		FS :	REAL := 5.0;
		LIMIT_L :	REAL;
		LIMIT_H :	REAL := 100.0;
		RST_VAL :	REAL;
		SET_VAL :	REAL := 100.0;
		TR :	TIME := T#500ms;
		S1 :	REAL := 2.0;
		S2 :	REAL := 10.0;
	END_VAR

	VAR_OUTPUT
		Y :	REAL;
	END_VAR

	VAR
		tx :	UDINT;
		start :	UDINT;
		state :	INT;
		in :	BOOL;
		step2 :	REAL;
		speed :	REAL;
		Y_start :	REAL;
		T_PLC_MS :	T_PLC_MS_block;
	END_VAR

	T_PLC_MS();
	tx:= T_PLC_MS.T_PLC_MS;

	IF rst THEN
		Y := RST_val;
		state := 0;
	ELSIF set THEN
		Y := SET_val;
		state := 0;
	ELSIF state > 0 THEN
		CASE state OF
			1 :
				in := su;
			2 :
				in := sd;
			3 :
				in := fu;
			4 :
				in := fd;
		END_CASE;
		IF NOT in AND tx - start <= TIME_TO_UDINT2(TR) THEN
			Y := Y_start + step2;
			state := 0;
		ELSIF in AND tx - start >= TIME_TO_UDINT2(TR) THEN
			Y := Y_start + UDINT_TO_REAL(tx - start - TIME_TO_UDINT2(TR)) * speed;
		ELSIF NOT in THEN
			state := 0;
		END_IF;
	ELSIF su THEN
		state := 1;
		start := tx;
		step2 := ss;
		speed := s1 * 1.0E-3;
		Y_start := Y;
	ELSIF sd THEN
		state := 2;
		start := tx;
		step2 := -ss;
		speed := -s1 * 1.0E-3;
		Y_start := Y;
	ELSIF fu THEN
		state := 3;
		start := tx;
		step2 := fs;
		speed := s2 * 1.0E-3;
		y_start := Y;
	ELSIF fd THEN
		state := 4;
		start := tx;
		step2 := -fs;
		speed := -s2 * 1.0E-3;
		y_start := Y;
	END_IF;
END_FUNCTION_BLOCK

PROGRAM program0
  	VAR
		SET :	BOOL;
		SU :	BOOL;
		SD :	BOOL;
		FU :	BOOL;
		FD :	BOOL;
		RST :	BOOL;
		SS :	REAL;
		FS :	REAL;
		LIMIT_L :	REAL;
		LIMIT_H :	REAL;
		RST_VAL :	REAL;
		SET_VAL :	REAL;
		TR :	TIME ;
		S1 :	REAL;
		S2 :	REAL;
		Y :	REAL;
		func_block : TUNE2_Block;
  	END_VAR
	func_block.SET := SET;
	func_block.SU := SU;
	func_block.SD := SD;
	func_block.FU := FU;
	func_block.FD := FD;
	func_block.RST := RST;
	func_block.SS:= SS;
	func_block.FS := FS;
	func_block.LIMIT_L := LIMIT_L;
	func_block.LIMIT_H := LIMIT_H;
	func_block.RST_VAL := RST_VAL;
	func_block.SET_VAL := SET_VAL;
	func_block.TR := TR;
	func_block.S1 := S1;
	func_block.S2 := S2;
	func_block();
	Y := func_block.Y;
END_PROGRAM

CONFIGURATION Config0
	VAR_GLOBAL
		PLC_TICKS_PER_SEC :	INT;
		PLC_SYS_TICK_CNT :	DINT;
	END_VAR

	RESOURCE Res0 ON PLC
		TASK task0(INTERVAL := T#20ms,PRIORITY := 0);
		PROGRAM instance0 WITH task0 : program0;
	END_RESOURCE
END_CONFIGURATION

(* ---- UPPERCASE.ST ---- *)
FUNCTION_BLOCK UPPERCASE_Block

	VAR_INPUT
		STR :	STRING;
	END_VAR

	VAR_OUTPUT
		UPPERCASE :	STRING;
	END_VAR

	VAR
		char :	BYTE;
		char2 :	BYTE;
		pos :	INT;
		l :	INT;
		str_temp :	STRING;
	END_VAR

	UPPERCASE := str;
	l := LEN(str);
	FOR pos := 1 TO l DO
		char := INT_TO_BYTE(GET_CHAR(str,pos));
		char2 := TO_UPPER(char);
		IF char <> char2 THEN
			str_temp := UPPERCASE;
			UPPERCASE := REPLACE(str_temp,BYTE_TO_STRING(char2,'%c'),1,pos);
		END_IF;
	END_FOR;

END_FUNCTION_BLOCK

PROGRAM program0
	VAR
	    LocalVar1 : STRING;
		LocalOUT  : STRING;
		func_block : UPPERCASE_Block;
  	END_VAR
	func_block.STR := LocalVar1;
	func_block();
	LocalOUT := func_block.UPPERCASE;
END_PROGRAM

CONFIGURATION Config0
  	RESOURCE Res0 ON PLC
    	TASK task0(INTERVAL := T#20ms,PRIORITY := 0);
    	PROGRAM instance0 WITH task0 : program0;
  	END_RESOURCE
END_CONFIGURATION

(* ---- URL_DECODE.ST ---- *)
TYPE
  oscat_STRING250               : STRING;
  oscat_STRING20               : STRING;
END_TYPE

FUNCTION_BLOCK HEX_TO_DWORD_Block

	VAR_INPUT
		HEX :	oscat_STRING20;
	END_VAR

	VAR_OUTPUT
		HEX_TO_DWORD :	DWORD;
	END_VAR

	VAR
		i :	INT;
		stop :	INT;
		X :	INT;
	END_VAR

	HEX_TO_DWORD := DWORD#0;
	stop := LEN(Hex);
	FOR I := 1 TO stop DO
		x := GET_CHAR(Hex,I);
		IF X > 47 AND x < 58 THEN
			HEX_TO_DWORD := SHL_DWORD(HEX_TO_DWORD,4) OR INT_TO_DWORD (X - 48);
		ELSIF X > 64 AND X < 71 THEN
			HEX_TO_DWORD := SHL_DWORD(HEX_TO_DWORD,4) OR INT_TO_DWORD (X - 55);
		ELSIF X > 96 AND X < 103 THEN
			HEX_TO_DWORD := SHL_DWORD(HEX_TO_DWORD,4) OR INT_TO_DWORD (X - 87);
		END_IF;
	END_FOR;

END_FUNCTION_BLOCK

FUNCTION_BLOCK URL_DECODE_Block

	VAR_INPUT
		IN :	oscat_STRING250;
	END_VAR

	VAR_OUTPUT
		URL_DECODE :	oscat_STRING250;
	END_VAR

	VAR
		pos :	INT;
		new :	STRING;
		HEX_TO_DWORD :	HEX_TO_DWORD_Block;
	END_VAR

	URL_DECODE := IN;
	pos := FIND(URL_DECODE,'%');
	WHILE pos > 0 DO
		HEX_TO_DWORD(Hex:=MID(URL_DECODE,2,pos + 1));
		new := BYTE_TO_STRING(DWORD_TO_BYTE(HEX_TO_DWORD.HEX_TO_DWORD),'%c');
		URL_DECODE := REPLACE(URL_DECODE, new, 3, pos);
		pos := FIND(URL_DECODE,'%');
	END_WHILE;

END_FUNCTION_BLOCK

PROGRAM program0
	VAR
		IN :	oscat_STRING250;
		URL_DECODE :	oscat_STRING250;

		func_block : URL_DECODE_Block;
	END_VAR
	func_block.IN := IN;

	func_block();
	URL_DECODE  := func_block.URL_DECODE;
END_PROGRAM

CONFIGURATION Config0
	RESOURCE Res0 ON PLC
		TASK task0(INTERVAL := T#20ms,PRIORITY := 0);
		PROGRAM instance0 WITH task0 : program0;
	END_RESOURCE
END_CONFIGURATION

(* ---- URL_ENCODE.ST ---- *)
FUNCTION_BLOCK URL_ENCODE_Block

	VAR_INPUT
		IN :	oscat_STRING250;
	END_VAR

	VAR_OUTPUT
		URL_ENCODE :	oscat_STRING250;
	END_VAR

	VAR
		pos_in :	INT;
		pos_out :	INT;
		stop :	INT;
		tb :	BYTE;
		pt_out :	oscat_aB1_255;
		char :	BYTE;
		BUF_TO_STRING :	BUF_TO_STRING;
		i :	INT;
	END_VAR

	pos_in := 1;
	stop := LEN(in);
	FOR pos_out := 1 TO 250 DO
		char := INT_TO_BYTE(GET_CHAR(IN,pos_in));
		IF pos_in > stop THEN
			EXIT;
		ELSIF IS_URLCHR(char) THEN
			pt_out[pos_out] := char;
			pos_in := pos_in + 1;
		ELSE
			IF pos_out > 248 THEN EXIT; END_IF;
			pt_out[pos_out] := BYTE#37;
			pos_out := pos_out + 1;
			tb := SHR_BYTE(char,4);
			IF tb > BYTE#9 THEN
				pt_out[pos_out] := USINT_TO_BYTE(BYTE_TO_USINT(tb) + USINT#55);
			ELSE
				pt_out[pos_out] := USINT_TO_BYTE(BYTE_TO_USINT(tb) + USINT#48);
			END_IF;
			pos_out := pos_out + 1;
			tb := char AND BYTE#16#0F;
			IF tb > BYTE#9 THEN
				pt_out[pos_out] := USINT_TO_BYTE(BYTE_TO_USINT(tb) + USINT#55);
			ELSE
				pt_out[pos_out] := USINT_TO_BYTE(BYTE_TO_USINT(tb) + USINT#48);
			END_IF;
			pos_in := pos_in + 1;
		END_IF;
	END_FOR;

	pos_out := pos_out - 1;

	FOR i := 0 TO 1 DO
	BUF_TO_STRING.REQ        := i>0;
	BUF_TO_STRING.BUF_FORMAT := TRUE;
	BUF_TO_STRING.BUF_OFFS   := DINT#0;
	BUF_TO_STRING.BUF_CNT    := INT_TO_DINT(pos_out);
	BUF_TO_STRING.BUFFER     := pt_out;
	BUF_TO_STRING.DST        := URL_ENCODE;
	BUF_TO_STRING();
	pt_out  := BUF_TO_STRING.BUFFER;
	URL_ENCODE := BUF_TO_STRING.DST;
	END_FOR;

END_FUNCTION_BLOCK

PROGRAM program0
	VAR
		IN :	oscat_STRING250;
		URL_ENCODE :	oscat_STRING250;

		func_block : URL_ENCODE_Block;
	END_VAR
	func_block.IN := IN;

	func_block();
	URL_ENCODE  := func_block.URL_ENCODE;
END_PROGRAM

CONFIGURATION Config0
	RESOURCE Res0 ON PLC
		TASK task0(INTERVAL := T#20ms,PRIORITY := 0);
		PROGRAM instance0 WITH task0 : program0;
	END_RESOURCE
END_CONFIGURATION

(* ---- URL_TO_STRING.ST ---- *)
TYPE
  oscat_STRING3               : STRING;
  oscat_STRING8               : STRING;
  oscat_STRING10              : STRING;
  oscat_STRING40              : STRING;
  oscat_STRING32              : STRING;
  oscat_STRING80              : STRING;
  oscat_STRING160              : STRING;
  oscat_STRING250              : STRING;
END_TYPE

TYPE oscat_url :
	STRUCT
		PROTOCOL : oscat_STRING10;
		USER     : oscat_STRING32;
		PASSWORD : oscat_STRING32;
		DOMAIN   : oscat_STRING80;
		PORT     : WORD;
		PATH     : oscat_STRING80;
		QUERY    : oscat_STRING250;
		ANCHOR   : oscat_STRING40;
		HEADER   : oscat_STRING160;
	END_STRUCT;
END_TYPE

FUNCTION_BLOCK URL_TO_STRING_Block

	VAR_INPUT
		IN :	oscat_url;
	END_VAR

	VAR_OUTPUT
		URL_TO_STRING :	oscat_STRING250;
	END_VAR

	IF NE_STRING(IN.PROTOCOL,'') THEN URL_TO_STRING := CONCAT(IN.PROTOCOL,'://'); END_IF;

	IF NE_STRING(IN.USER,'') THEN
		URL_TO_STRING := CONCAT(URL_TO_STRING, IN.USER);
		IF NE_STRING(IN.PASSWORD,'') THEN
			URL_TO_STRING := CONCAT(URL_TO_STRING, ':');
			URL_TO_STRING := CONCAT(URL_TO_STRING, IN.PASSWORD);
		END_IF;
		URL_TO_STRING := CONCAT(URL_TO_STRING, '@');
	END_IF;

	URL_TO_STRING := CONCAT(URL_TO_STRING, IN.DOMAIN);

	IF IN.PORT > WORD#0 THEN
		URL_TO_STRING := CONCAT(URL_TO_STRING, ':');
		URL_TO_STRING := CONCAT(URL_TO_STRING, WORD_TO_STRING(IN.PORT));
	END_IF;

	URL_TO_STRING := CONCAT(URL_TO_STRING, IN.PATH);

	IF NE_STRING(IN.QUERY,'') THEN
		URL_TO_STRING := CONCAT(URL_TO_STRING, '?');
		URL_TO_STRING := CONCAT(URL_TO_STRING, IN.QUERY);
	END_IF;

	IF NE_STRING(IN.ANCHOR,'') THEN
		URL_TO_STRING := CONCAT(URL_TO_STRING, '#');
		URL_TO_STRING := CONCAT(URL_TO_STRING, IN.ANCHOR);
	END_IF;

END_FUNCTION_BLOCK

PROGRAM program0
	VAR
		IN :	oscat_url;
		URL_TO_STRING :	oscat_STRING250;

		func_block : URL_TO_STRING_Block;
	END_VAR
	func_block.IN := IN;

	func_block();
	URL_TO_STRING  := func_block.URL_TO_STRING;
END_PROGRAM

CONFIGURATION Config0
	RESOURCE Res0 ON PLC
		TASK task0(INTERVAL := T#20ms,PRIORITY := 0);
		PROGRAM instance0 WITH task0 : program0;
	END_RESOURCE
END_CONFIGURATION

(* ---- V3_ABS.ST ---- *)
TYPE oscat_vector_3:
	STRUCT
		X : REAL;
		Y : REAL;
		Z : REAL;
	END_STRUCT;
END_TYPE

FUNCTION_BLOCK V3_ABS_Block

	VAR_INPUT
		A :	oscat_vector_3;
	END_VAR

	VAR_OUTPUT
		V3_ABS :	REAL;
	END_VAR

	V3_ABS := SQRT(A.X * A.X + A.Y * A.Y + A.Z * A.Z);

END_FUNCTION_BLOCK

PROGRAM program0
  	VAR
		A :	oscat_vector_3;
		V3_ABS :	REAL;
		func_block : V3_ABS_Block;
  	END_VAR
	func_block.A := A;
	func_block();
	V3_ABS := func_block.V3_ABS;
END_PROGRAM

CONFIGURATION Config0
	RESOURCE Res0 ON PLC
		TASK task0(INTERVAL := T#20ms,PRIORITY := 0);
		PROGRAM instance0 WITH task0 : program0;
	END_RESOURCE
END_CONFIGURATION

(* ---- V3_ADD.ST ---- *)
TYPE oscat_vector_3:
	STRUCT
		X : REAL;
		Y : REAL;
		Z : REAL;
	END_STRUCT;
END_TYPE

FUNCTION_BLOCK V3_ADD_Block
	VAR_INPUT
		A :	oscat_vector_3;
		B :	oscat_vector_3;
	END_VAR

	VAR_OUTPUT
		V3_ADD :	oscat_vector_3;
	END_VAR

	V3_ADD.X := A.X + B.X;
	V3_ADD.Y := A.Y + B.Y;
	V3_ADD.Z := A.Z + B.Z;

END_FUNCTION_BLOCK

PROGRAM program0
  	VAR
		A :	oscat_vector_3;
		B :	oscat_vector_3;
		V3_ADD :	oscat_vector_3;
		func_block : V3_ADD_Block;
  	END_VAR
	func_block.A := A;
	func_block.B := B;
	func_block();
	V3_ADD := func_block.V3_ADD;
END_PROGRAM

CONFIGURATION Config0
  RESOURCE Res0 ON PLC
    TASK task0(INTERVAL := T#20ms,PRIORITY := 0);
    PROGRAM instance0 WITH task0 : program0;
  END_RESOURCE
END_CONFIGURATION

(* ---- V3_ANG.ST ---- *)
TYPE oscat_vector_3:
	STRUCT
		X : REAL;
		Y : REAL;
		Z : REAL;
	END_STRUCT;
END_TYPE

FUNCTION_BLOCK V3_ABS_Block
	VAR_INPUT
		A :	oscat_vector_3;
	END_VAR

	VAR_OUTPUT
		V3_ABS : REAL;
	END_VAR

	V3_ABS := SQRT(A.X * A.X + A.Y * A.Y + A.Z * A.Z);

END_FUNCTION_BLOCK

FUNCTION_BLOCK V3_DPRO_Block

	VAR_INPUT
		A :	oscat_vector_3;
		B :	oscat_vector_3;
	END_VAR

	VAR_OUTPUT
		V3_DPRO :	REAL;
	END_VAR

	V3_DPRO := A.X * B.X + A.Y * B.Y + A.Z * B.Z;

END_FUNCTION_BLOCK

FUNCTION_BLOCK V3_ANG_Block

	VAR_INPUT
		A :	oscat_vector_3;
		B :	oscat_vector_3;
	END_VAR

	VAR_OUTPUT
		V3_ANG :	REAL;
	END_VAR

	VAR
		d :	REAL;
		V3_ABS :	V3_ABS_Block;
		V3_DPRO :	V3_DPRO_Block;
	END_VAR

	V3_ABS(A:=A);
	d :=V3_ABS.V3_ABS;

	V3_ABS(A:=B);
	d := d * V3_ABS.V3_ABS;

	IF d > 0.0 THEN
		V3_DPRO(A:=A,B:=B);
		V3_ANG := ACOS(LIMIT(-1.0, V3_DPRO.V3_DPRO / d,1.0));
	ELSE
		V3_ANG := 0.0;

	END_IF;

END_FUNCTION_BLOCK

PROGRAM program0
  	VAR
		A :	oscat_vector_3;
		B :	oscat_vector_3;
		V3_ANG :	REAL;
		func_block : V3_ANG_Block;
  	END_VAR
	func_block.A := A;
	func_block.B := B;
	func_block();
	V3_ANG := func_block.V3_ANG;
END_PROGRAM

CONFIGURATION Config0
  RESOURCE Res0 ON PLC
    TASK task0(INTERVAL := T#20ms,PRIORITY := 0);
    PROGRAM instance0 WITH task0 : program0;
  END_RESOURCE
END_CONFIGURATION

(* ---- V3_DPRO.ST ---- *)
TYPE oscat_vector_3:
	STRUCT
		X : REAL;
		Y : REAL;
		Z : REAL;
	END_STRUCT;
END_TYPE

FUNCTION_BLOCK V3_DPRO_Block

	VAR_INPUT
		A :	oscat_vector_3;
		B :	oscat_vector_3;
	END_VAR

	VAR_OUTPUT
		V3_DPRO :	REAL;
	END_VAR

	V3_DPRO := A.X * B.X + A.Y * B.Y + A.Z * B.Z;

END_FUNCTION_BLOCK

PROGRAM program0
  	VAR
		A :	oscat_vector_3;
		B :	oscat_vector_3;
		V3_DPRO : REAL;
		func_block : V3_DPRO_Block;
  	END_VAR
	func_block.A := A;
	func_block.B := B;
	func_block();
	V3_DPRO := func_block.V3_DPRO;
END_PROGRAM

CONFIGURATION Config0
  RESOURCE Res0 ON PLC
    TASK task0(INTERVAL := T#20ms,PRIORITY := 0);
    PROGRAM instance0 WITH task0 : program0;
  END_RESOURCE
END_CONFIGURATION

(* ---- V3_NORM.ST ---- *)
TYPE oscat_vector_3:
	STRUCT
		X : REAL;
		Y : REAL;
		Z : REAL;
	END_STRUCT;
END_TYPE

FUNCTION_BLOCK V3_ABS_Block

	VAR_INPUT
		A :	oscat_vector_3;
	END_VAR

	VAR_OUTPUT
		V3_ABS :	REAL;
	END_VAR

	V3_ABS := SQRT(A.X * A.X + A.Y * A.Y + A.Z * A.Z);

END_FUNCTION_BLOCK

FUNCTION_BLOCK V3_SMUL_Block
	VAR_INPUT
		A :	oscat_vector_3;
		M :	REAL;
	END_VAR

	VAR_OUTPUT
		V3_SMUL :	oscat_vector_3;
	END_VAR

	V3_SMUL.X := A.X * M;
	V3_SMUL.Y := A.Y * M;
	V3_SMUL.Z := A.Z * M;
END_FUNCTION_BLOCK

FUNCTION_BLOCK V3_NORM_Block

	VAR_INPUT
		A :	oscat_vector_3;
	END_VAR

	VAR_OUTPUT
		V3_NORM :	oscat_vector_3;
	END_VAR

	VAR
		la :	REAL;
		V3_SMUL :	V3_SMUL_Block;
		V3_ABS :	V3_ABS_Block;
	END_VAR

	V3_ABS(A:=A);
	la:=V3_ABS.V3_ABS;

	IF la > 0.0 THEN
		V3_SMUL(A:=A,M:=1.0/la);
		V3_NORM:=V3_SMUL.V3_SMUL;
	ELSE
		V3_NORM.X := 0.0;
		V3_NORM.Y := 0.0;
		V3_NORM.Z := 0.0;
	END_IF;

END_FUNCTION_BLOCK

PROGRAM program0
  	VAR
		A :	oscat_vector_3;
		V3_NORM :	oscat_vector_3;
		func_block : V3_NORM_Block;
  	END_VAR
	func_block.A := A;
	func_block();
	V3_NORM := func_block.V3_NORM;
END_PROGRAM

CONFIGURATION Config0
  RESOURCE Res0 ON PLC
    TASK task0(INTERVAL := T#20ms,PRIORITY := 0);
    PROGRAM instance0 WITH task0 : program0;
  END_RESOURCE
END_CONFIGURATION

(* ---- V3_NUL.ST ---- *)
TYPE oscat_vector_3:
	STRUCT
		X : REAL;
		Y : REAL;
		Z : REAL;
	END_STRUCT;
END_TYPE

FUNCTION_BLOCK V3_NUL_Block

	VAR_INPUT
		A :	oscat_vector_3;
	END_VAR

	VAR_OUTPUT
		V3_NUL :	BOOL;
	END_VAR

	V3_NUL := A.X = 0.0 AND A.Y = 0.0 AND A.Z = 0.0;

END_FUNCTION_BLOCK

PROGRAM program0
  	VAR
		A :	oscat_vector_3;
		V3_NUL :	BOOL;
		func_block : V3_NUL_Block;
  	END_VAR
	func_block.A := A;
	func_block();
	V3_NUL := func_block.V3_NUL;
END_PROGRAM

CONFIGURATION Config0
  RESOURCE Res0 ON PLC
    TASK task0(INTERVAL := T#20ms,PRIORITY := 0);
    PROGRAM instance0 WITH task0 : program0;
  END_RESOURCE
END_CONFIGURATION

(* ---- V3_PAR.ST ---- *)
TYPE oscat_vector_3:
	STRUCT
		X : REAL;
		Y : REAL;
		Z : REAL;
	END_STRUCT;
END_TYPE

FUNCTION_BLOCK V3_ABS_Block

	VAR_INPUT
		A :	oscat_vector_3;
	END_VAR

	VAR_OUTPUT
		V3_ABS :	REAL;
	END_VAR

	V3_ABS := SQRT(A.X * A.X + A.Y * A.Y + A.Z * A.Z);

END_FUNCTION_BLOCK

FUNCTION_BLOCK V3_XPRO_Block
	VAR_INPUT
		A :	oscat_vector_3;
		B :	oscat_vector_3;
	END_VAR

	VAR_OUTPUT
		V3_XPRO :	oscat_vector_3;
	END_VAR

	V3_XPRO.X := A.Y * B.Z - A.Z * B.Y;
	V3_XPRO.Y := A.Z * B.X - A.X * B.Z;
	V3_XPRO.Z := A.X * B.Y - A.Y * B.X;

END_FUNCTION_BLOCK

FUNCTION_BLOCK V3_PAR_Block
	VAR_INPUT
		A :	oscat_vector_3;
		B :	oscat_vector_3;
	END_VAR

	VAR_OUTPUT
		V3_PAR :	BOOL;
	END_VAR

	VAR
		V3_XPRO :	V3_XPRO_Block;
		V3_ABS :	V3_ABS_Block;
	END_VAR

	V3_XPRO(A:=A,B:=B);
	V3_ABS(A:=V3_XPRO.V3_XPRO);

	V3_PAR := V3_ABS.V3_ABS = 0.0;

END_FUNCTION_BLOCK

PROGRAM program0
  	VAR
		A :	oscat_vector_3;
		B :	oscat_vector_3;
		V3_PAR :	BOOL;
		func_block : V3_PAR_Block;
  	END_VAR
	func_block.A := A;
	func_block.B := B;
	func_block();
	V3_PAR := func_block.V3_PAR;
END_PROGRAM

CONFIGURATION Config0
  RESOURCE Res0 ON PLC
    TASK task0(INTERVAL := T#20ms,PRIORITY := 0);
    PROGRAM instance0 WITH task0 : program0;
  END_RESOURCE
END_CONFIGURATION

(* ---- V3_REV.ST ---- *)
TYPE oscat_vector_3:
	STRUCT
		X : REAL;
		Y : REAL;
		Z : REAL;
	END_STRUCT;
END_TYPE

FUNCTION_BLOCK V3_REV_Block
	VAR_INPUT
		A :	oscat_vector_3;
	END_VAR

	VAR_OUTPUT
		V3_REV :	oscat_vector_3;
	END_VAR

	V3_REV.X := -A.X;
	V3_REV.Y := -A.Y;
	V3_REV.Z := -A.Z;

END_FUNCTION_BLOCK

PROGRAM program0
  	VAR
		A :	oscat_vector_3;
		V3_REV : oscat_vector_3;
		func_block : V3_REV_Block;
  	END_VAR
	func_block.A := A;
	func_block();
	V3_REV := func_block.V3_REV;
END_PROGRAM

CONFIGURATION Config0
  RESOURCE Res0 ON PLC
    TASK task0(INTERVAL := T#20ms,PRIORITY := 0);
    PROGRAM instance0 WITH task0 : program0;
  END_RESOURCE
END_CONFIGURATION

(* ---- V3_SMUL.ST ---- *)
TYPE oscat_vector_3:
	STRUCT
		X : REAL;
		Y : REAL;
		Z : REAL;
	END_STRUCT;
END_TYPE

FUNCTION_BLOCK V3_SMUL_Block
	VAR_INPUT
		A :	oscat_vector_3;
		M :	REAL;
	END_VAR

	VAR_OUTPUT
		V3_SMUL :	oscat_vector_3;
	END_VAR

	V3_SMUL.X := A.X * M;
	V3_SMUL.Y := A.Y * M;
	V3_SMUL.Z := A.Z * M;
END_FUNCTION_BLOCK

PROGRAM program0
  	VAR
		A :	oscat_vector_3;
		M :	REAL;
		V3_SMUL :	oscat_vector_3;
		func_block : V3_SMUL_Block;
  	END_VAR
	func_block.A := A;
	func_block.M := M;
	func_block();
	V3_SMUL := func_block.V3_SMUL;
END_PROGRAM

CONFIGURATION Config0
	RESOURCE Res0 ON PLC
		TASK task0(INTERVAL := T#20ms,PRIORITY := 0);
		PROGRAM instance0 WITH task0 : program0;
	END_RESOURCE
END_CONFIGURATION

(* ---- V3_SUB.ST ---- *)
TYPE oscat_vector_3:
	STRUCT
		X : REAL;
		Y : REAL;
		Z : REAL;
	END_STRUCT;
END_TYPE

FUNCTION_BLOCK V3_SUB_Block

	VAR_INPUT
		A :	oscat_vector_3;
		B :	oscat_vector_3;
	END_VAR

	VAR_OUTPUT
		V3_SUB :	oscat_vector_3;
	END_VAR

	V3_SUB.X := A.X - B.X;
	V3_SUB.Y := A.Y - B.Y;
	V3_SUB.Z := A.Z - B.Z;

END_FUNCTION_BLOCK

PROGRAM program0
  	VAR
		A :	oscat_vector_3;
		B :	oscat_vector_3;
		V3_SUB :	oscat_vector_3;
		func_block : V3_SUB_Block;
  	END_VAR
	func_block.A := A;
	func_block.B := B;
	func_block();
	V3_SUB := func_block.V3_SUB;
END_PROGRAM

CONFIGURATION Config0
  RESOURCE Res0 ON PLC
    TASK task0(INTERVAL := T#20ms,PRIORITY := 0);
    PROGRAM instance0 WITH task0 : program0;
  END_RESOURCE
END_CONFIGURATION

(* ---- V3_XANG.ST ---- *)
TYPE oscat_vector_3 :
	STRUCT
		X : REAL;
		Y : REAL;
		Z : REAL;
	END_STRUCT;
END_TYPE

FUNCTION_BLOCK V3_ABS_Block

	VAR_INPUT
		A :	oscat_vector_3;
	END_VAR

	VAR_OUTPUT
		V3_ABS :	REAL;
	END_VAR

	V3_ABS := SQRT(A.X * A.X + A.Y * A.Y + A.Z * A.Z);

END_FUNCTION_BLOCK

FUNCTION_BLOCK V3_XANG_Block

	VAR_INPUT
		A :	oscat_vector_3;
	END_VAR

	VAR_OUTPUT
		V3_XANG :	REAL;
	END_VAR

	VAR
		la :	REAL;
		V3_ABS :	V3_ABS_Block;
	END_VAR

	V3_ABS(A:=A);
	la:=V3_ABS.V3_ABS;

	IF la > 0.0 THEN
		V3_XANG := ACOS(A.X / la);
	ELSE
		V3_XANG := 0.0;
	END_IF;

END_FUNCTION_BLOCK

PROGRAM program0
  	VAR
		A :	oscat_vector_3;
		V3_XANG :	REAL;
		func_block : V3_XANG_Block;
  	END_VAR
	func_block.A := A;
	func_block();
	V3_XANG := func_block.V3_XANG;
END_PROGRAM

CONFIGURATION Config0
  RESOURCE Res0 ON PLC
    TASK task0(INTERVAL := T#20ms,PRIORITY := 0);
    PROGRAM instance0 WITH task0 : program0;
  END_RESOURCE
END_CONFIGURATION
